(* IEC 61131-3 sources: 2026_Projet_YGO_ExcavatriceDragage/TOOLS/TEST_AUTO_CI/RESULTS/L_SIMULATION/tests (part 10) *)

TEST 'TC-T418-INT-009 Reference etablie N1 puis cycle sans depart homing'
nx := 5000; ny := 5000; raw1 := 0; raw2 := 0; previousButton := FALSE; buttonEdges := 0;
bench.Enable := TRUE; joy.Enable := TRUE; joy.ArmingPermit := TRUE; diagOk.Operational := TRUE; joy.BusCanOpenOP := diagOk; joy.JoystickOP := diagOk;
home.Enable := TRUE; home.BootReady := TRUE; home.Mode := E_Mode.MAINT_N1; home.WinchesMechanicallyStopped := TRUE;
(* Fixture deja referencee : les preuves du preset manuel reel sont dans la CI codeurs/benne et le routage PRG inchange. *)
home.M1Status.HomedAndReliable := TRUE; home.M2Status.HomedAndReliable := TRUE; home.BucketOffsetValid := TRUE;
ADVANCE_TIME(10000000); bench(RawPosM1 := raw1, RawPosM2 := raw2);
joy(RawX := bench.Operator.JoyXRaw_ANA1, RawY := bench.Operator.JoyYRaw_ANA2, RawButton := bench.Operator.JoyBtnRaw, Cfg := cfg, NeutralXMem := nx, NeutralYMem := ny);
home(DeadmanArmed := joy.DeadmanArmed, JoystickDeflected := NOT joy.AtNeutralXY, JoystickPull := joy.AxisCmdY.DirectionPositive, JoystickPush := joy.AxisCmdY.DirectionNegative, BtnValidation := bench.Operator.JoyBtnRaw);
ASSERT_EQ(home.MachineHomingSeqStep, E_MachineHomingTxState.HX0_REPOS, 'N1/cycle : aucun HX1 par geste joystick'); ASSERT_FALSE(home.M3Locked, 'N1/cycle : aucun verrou homing parasite'); ASSERT_TRUE(home.MachineHomed, 'Reference conservee');
bench.SimJoystickFwd_Up_Close_Active := TRUE;
ADVANCE_TIME(10000000); bench(RawPosM1 := raw1, RawPosM2 := raw2);
joy(RawX := bench.Operator.JoyXRaw_ANA1, RawY := bench.Operator.JoyYRaw_ANA2, RawButton := bench.Operator.JoyBtnRaw, Cfg := cfg, NeutralXMem := nx, NeutralYMem := ny);
home(DeadmanArmed := joy.DeadmanArmed, JoystickDeflected := NOT joy.AtNeutralXY, JoystickPull := joy.AxisCmdY.DirectionPositive, JoystickPush := joy.AxisCmdY.DirectionNegative, BtnValidation := bench.Operator.JoyBtnRaw);
ASSERT_EQ(home.MachineHomingSeqStep, E_MachineHomingTxState.HX0_REPOS, 'N1/cycle : aucun HX1 par geste joystick'); ASSERT_FALSE(home.M3Locked, 'N1/cycle : aucun verrou homing parasite'); ASSERT_TRUE(home.MachineHomed, 'Reference conservee');
ADVANCE_TIME(10000000); bench(RawPosM1 := raw1, RawPosM2 := raw2);
joy(RawX := bench.Operator.JoyXRaw_ANA1, RawY := bench.Operator.JoyYRaw_ANA2, RawButton := bench.Operator.JoyBtnRaw, Cfg := cfg, NeutralXMem := nx, NeutralYMem := ny);
home(DeadmanArmed := joy.DeadmanArmed, JoystickDeflected := NOT joy.AtNeutralXY, JoystickPull := joy.AxisCmdY.DirectionPositive, JoystickPush := joy.AxisCmdY.DirectionNegative, BtnValidation := bench.Operator.JoyBtnRaw);
ASSERT_EQ(home.MachineHomingSeqStep, E_MachineHomingTxState.HX0_REPOS, 'N1/cycle : aucun HX1 par geste joystick'); ASSERT_FALSE(home.M3Locked, 'N1/cycle : aucun verrou homing parasite'); ASSERT_TRUE(home.MachineHomed, 'Reference conservee');
ADVANCE_TIME(10000000); bench(RawPosM1 := raw1, RawPosM2 := raw2);
joy(RawX := bench.Operator.JoyXRaw_ANA1, RawY := bench.Operator.JoyYRaw_ANA2, RawButton := bench.Operator.JoyBtnRaw, Cfg := cfg, NeutralXMem := nx, NeutralYMem := ny);
home(DeadmanArmed := joy.DeadmanArmed, JoystickDeflected := NOT joy.AtNeutralXY, JoystickPull := joy.AxisCmdY.DirectionPositive, JoystickPush := joy.AxisCmdY.DirectionNegative, BtnValidation := bench.Operator.JoyBtnRaw);
ASSERT_EQ(home.MachineHomingSeqStep, E_MachineHomingTxState.HX0_REPOS, 'N1/cycle : aucun HX1 par geste joystick'); ASSERT_FALSE(home.M3Locked, 'N1/cycle : aucun verrou homing parasite'); ASSERT_TRUE(home.MachineHomed, 'Reference conservee');
ADVANCE_TIME(10000000); bench(RawPosM1 := raw1, RawPosM2 := raw2);
joy(RawX := bench.Operator.JoyXRaw_ANA1, RawY := bench.Operator.JoyYRaw_ANA2, RawButton := bench.Operator.JoyBtnRaw, Cfg := cfg, NeutralXMem := nx, NeutralYMem := ny);
home(DeadmanArmed := joy.DeadmanArmed, JoystickDeflected := NOT joy.AtNeutralXY, JoystickPull := joy.AxisCmdY.DirectionPositive, JoystickPush := joy.AxisCmdY.DirectionNegative, BtnValidation := bench.Operator.JoyBtnRaw);
ASSERT_EQ(home.MachineHomingSeqStep, E_MachineHomingTxState.HX0_REPOS, 'N1/cycle : aucun HX1 par geste joystick'); ASSERT_FALSE(home.M3Locked, 'N1/cycle : aucun verrou homing parasite'); ASSERT_TRUE(home.MachineHomed, 'Reference conservee');
ADVANCE_TIME(10000000); bench(RawPosM1 := raw1, RawPosM2 := raw2);
joy(RawX := bench.Operator.JoyXRaw_ANA1, RawY := bench.Operator.JoyYRaw_ANA2, RawButton := bench.Operator.JoyBtnRaw, Cfg := cfg, NeutralXMem := nx, NeutralYMem := ny);
home(DeadmanArmed := joy.DeadmanArmed, JoystickDeflected := NOT joy.AtNeutralXY, JoystickPull := joy.AxisCmdY.DirectionPositive, JoystickPush := joy.AxisCmdY.DirectionNegative, BtnValidation := bench.Operator.JoyBtnRaw);
ASSERT_EQ(home.MachineHomingSeqStep, E_MachineHomingTxState.HX0_REPOS, 'N1/cycle : aucun HX1 par geste joystick'); ASSERT_FALSE(home.M3Locked, 'N1/cycle : aucun verrou homing parasite'); ASSERT_TRUE(home.MachineHomed, 'Reference conservee');
ADVANCE_TIME(10000000); bench(RawPosM1 := raw1, RawPosM2 := raw2);
joy(RawX := bench.Operator.JoyXRaw_ANA1, RawY := bench.Operator.JoyYRaw_ANA2, RawButton := bench.Operator.JoyBtnRaw, Cfg := cfg, NeutralXMem := nx, NeutralYMem := ny);
home(DeadmanArmed := joy.DeadmanArmed, JoystickDeflected := NOT joy.AtNeutralXY, JoystickPull := joy.AxisCmdY.DirectionPositive, JoystickPush := joy.AxisCmdY.DirectionNegative, BtnValidation := bench.Operator.JoyBtnRaw);
ASSERT_EQ(home.MachineHomingSeqStep, E_MachineHomingTxState.HX0_REPOS, 'N1/cycle : aucun HX1 par geste joystick'); ASSERT_FALSE(home.M3Locked, 'N1/cycle : aucun verrou homing parasite'); ASSERT_TRUE(home.MachineHomed, 'Reference conservee');
ADVANCE_TIME(10000000); bench(RawPosM1 := raw1, RawPosM2 := raw2);
joy(RawX := bench.Operator.JoyXRaw_ANA1, RawY := bench.Operator.JoyYRaw_ANA2, RawButton := bench.Operator.JoyBtnRaw, Cfg := cfg, NeutralXMem := nx, NeutralYMem := ny);
home(DeadmanArmed := joy.DeadmanArmed, JoystickDeflected := NOT joy.AtNeutralXY, JoystickPull := joy.AxisCmdY.DirectionPositive, JoystickPush := joy.AxisCmdY.DirectionNegative, BtnValidation := bench.Operator.JoyBtnRaw);
ASSERT_EQ(home.MachineHomingSeqStep, E_MachineHomingTxState.HX0_REPOS, 'N1/cycle : aucun HX1 par geste joystick'); ASSERT_FALSE(home.M3Locked, 'N1/cycle : aucun verrou homing parasite'); ASSERT_TRUE(home.MachineHomed, 'Reference conservee');
ADVANCE_TIME(10000000); bench(RawPosM1 := raw1, RawPosM2 := raw2);
joy(RawX := bench.Operator.JoyXRaw_ANA1, RawY := bench.Operator.JoyYRaw_ANA2, RawButton := bench.Operator.JoyBtnRaw, Cfg := cfg, NeutralXMem := nx, NeutralYMem := ny);
home(DeadmanArmed := joy.DeadmanArmed, JoystickDeflected := NOT joy.AtNeutralXY, JoystickPull := joy.AxisCmdY.DirectionPositive, JoystickPush := joy.AxisCmdY.DirectionNegative, BtnValidation := bench.Operator.JoyBtnRaw);
ASSERT_EQ(home.MachineHomingSeqStep, E_MachineHomingTxState.HX0_REPOS, 'N1/cycle : aucun HX1 par geste joystick'); ASSERT_FALSE(home.M3Locked, 'N1/cycle : aucun verrou homing parasite'); ASSERT_TRUE(home.MachineHomed, 'Reference conservee');
ADVANCE_TIME(10000000); bench(RawPosM1 := raw1, RawPosM2 := raw2);
joy(RawX := bench.Operator.JoyXRaw_ANA1, RawY := bench.Operator.JoyYRaw_ANA2, RawButton := bench.Operator.JoyBtnRaw, Cfg := cfg, NeutralXMem := nx, NeutralYMem := ny);
home(DeadmanArmed := joy.DeadmanArmed, JoystickDeflected := NOT joy.AtNeutralXY, JoystickPull := joy.AxisCmdY.DirectionPositive, JoystickPush := joy.AxisCmdY.DirectionNegative, BtnValidation := bench.Operator.JoyBtnRaw);
ASSERT_EQ(home.MachineHomingSeqStep, E_MachineHomingTxState.HX0_REPOS, 'N1/cycle : aucun HX1 par geste joystick'); ASSERT_FALSE(home.M3Locked, 'N1/cycle : aucun verrou homing parasite'); ASSERT_TRUE(home.MachineHomed, 'Reference conservee');
ADVANCE_TIME(10000000); bench(RawPosM1 := raw1, RawPosM2 := raw2);
joy(RawX := bench.Operator.JoyXRaw_ANA1, RawY := bench.Operator.JoyYRaw_ANA2, RawButton := bench.Operator.JoyBtnRaw, Cfg := cfg, NeutralXMem := nx, NeutralYMem := ny);
home(DeadmanArmed := joy.DeadmanArmed, JoystickDeflected := NOT joy.AtNeutralXY, JoystickPull := joy.AxisCmdY.DirectionPositive, JoystickPush := joy.AxisCmdY.DirectionNegative, BtnValidation := bench.Operator.JoyBtnRaw);
ASSERT_EQ(home.MachineHomingSeqStep, E_MachineHomingTxState.HX0_REPOS, 'N1/cycle : aucun HX1 par geste joystick'); ASSERT_FALSE(home.M3Locked, 'N1/cycle : aucun verrou homing parasite'); ASSERT_TRUE(home.MachineHomed, 'Reference conservee');
ADVANCE_TIME(10000000); bench(RawPosM1 := raw1, RawPosM2 := raw2);
joy(RawX := bench.Operator.JoyXRaw_ANA1, RawY := bench.Operator.JoyYRaw_ANA2, RawButton := bench.Operator.JoyBtnRaw, Cfg := cfg, NeutralXMem := nx, NeutralYMem := ny);
home(DeadmanArmed := joy.DeadmanArmed, JoystickDeflected := NOT joy.AtNeutralXY, JoystickPull := joy.AxisCmdY.DirectionPositive, JoystickPush := joy.AxisCmdY.DirectionNegative, BtnValidation := bench.Operator.JoyBtnRaw);
ASSERT_EQ(home.MachineHomingSeqStep, E_MachineHomingTxState.HX0_REPOS, 'N1/cycle : aucun HX1 par geste joystick'); ASSERT_FALSE(home.M3Locked, 'N1/cycle : aucun verrou homing parasite'); ASSERT_TRUE(home.MachineHomed, 'Reference conservee');
ADVANCE_TIME(10000000); bench(RawPosM1 := raw1, RawPosM2 := raw2);
joy(RawX := bench.Operator.JoyXRaw_ANA1, RawY := bench.Operator.JoyYRaw_ANA2, RawButton := bench.Operator.JoyBtnRaw, Cfg := cfg, NeutralXMem := nx, NeutralYMem := ny);
home(DeadmanArmed := joy.DeadmanArmed, JoystickDeflected := NOT joy.AtNeutralXY, JoystickPull := joy.AxisCmdY.DirectionPositive, JoystickPush := joy.AxisCmdY.DirectionNegative, BtnValidation := bench.Operator.JoyBtnRaw);
ASSERT_EQ(home.MachineHomingSeqStep, E_MachineHomingTxState.HX0_REPOS, 'N1/cycle : aucun HX1 par geste joystick'); ASSERT_FALSE(home.M3Locked, 'N1/cycle : aucun verrou homing parasite'); ASSERT_TRUE(home.MachineHomed, 'Reference conservee');
ADVANCE_TIME(10000000); bench(RawPosM1 := raw1, RawPosM2 := raw2);
joy(RawX := bench.Operator.JoyXRaw_ANA1, RawY := bench.Operator.JoyYRaw_ANA2, RawButton := bench.Operator.JoyBtnRaw, Cfg := cfg, NeutralXMem := nx, NeutralYMem := ny);
home(DeadmanArmed := joy.DeadmanArmed, JoystickDeflected := NOT joy.AtNeutralXY, JoystickPull := joy.AxisCmdY.DirectionPositive, JoystickPush := joy.AxisCmdY.DirectionNegative, BtnValidation := bench.Operator.JoyBtnRaw);
ASSERT_EQ(home.MachineHomingSeqStep, E_MachineHomingTxState.HX0_REPOS, 'N1/cycle : aucun HX1 par geste joystick'); ASSERT_FALSE(home.M3Locked, 'N1/cycle : aucun verrou homing parasite'); ASSERT_TRUE(home.MachineHomed, 'Reference conservee');
ADVANCE_TIME(10000000); bench(RawPosM1 := raw1, RawPosM2 := raw2);
joy(RawX := bench.Operator.JoyXRaw_ANA1, RawY := bench.Operator.JoyYRaw_ANA2, RawButton := bench.Operator.JoyBtnRaw, Cfg := cfg, NeutralXMem := nx, NeutralYMem := ny);
home(DeadmanArmed := joy.DeadmanArmed, JoystickDeflected := NOT joy.AtNeutralXY, JoystickPull := joy.AxisCmdY.DirectionPositive, JoystickPush := joy.AxisCmdY.DirectionNegative, BtnValidation := bench.Operator.JoyBtnRaw);
ASSERT_EQ(home.MachineHomingSeqStep, E_MachineHomingTxState.HX0_REPOS, 'N1/cycle : aucun HX1 par geste joystick'); ASSERT_FALSE(home.M3Locked, 'N1/cycle : aucun verrou homing parasite'); ASSERT_TRUE(home.MachineHomed, 'Reference conservee');
ADVANCE_TIME(10000000); bench(RawPosM1 := raw1, RawPosM2 := raw2);
joy(RawX := bench.Operator.JoyXRaw_ANA1, RawY := bench.Operator.JoyYRaw_ANA2, RawButton := bench.Operator.JoyBtnRaw, Cfg := cfg, NeutralXMem := nx, NeutralYMem := ny);
home(DeadmanArmed := joy.DeadmanArmed, JoystickDeflected := NOT joy.AtNeutralXY, JoystickPull := joy.AxisCmdY.DirectionPositive, JoystickPush := joy.AxisCmdY.DirectionNegative, BtnValidation := bench.Operator.JoyBtnRaw);
ASSERT_EQ(home.MachineHomingSeqStep, E_MachineHomingTxState.HX0_REPOS, 'N1/cycle : aucun HX1 par geste joystick'); ASSERT_FALSE(home.M3Locked, 'N1/cycle : aucun verrou homing parasite'); ASSERT_TRUE(home.MachineHomed, 'Reference conservee');
ADVANCE_TIME(10000000); bench(RawPosM1 := raw1, RawPosM2 := raw2);
joy(RawX := bench.Operator.JoyXRaw_ANA1, RawY := bench.Operator.JoyYRaw_ANA2, RawButton := bench.Operator.JoyBtnRaw, Cfg := cfg, NeutralXMem := nx, NeutralYMem := ny);
home(DeadmanArmed := joy.DeadmanArmed, JoystickDeflected := NOT joy.AtNeutralXY, JoystickPull := joy.AxisCmdY.DirectionPositive, JoystickPush := joy.AxisCmdY.DirectionNegative, BtnValidation := bench.Operator.JoyBtnRaw);
ASSERT_EQ(home.MachineHomingSeqStep, E_MachineHomingTxState.HX0_REPOS, 'N1/cycle : aucun HX1 par geste joystick'); ASSERT_FALSE(home.M3Locked, 'N1/cycle : aucun verrou homing parasite'); ASSERT_TRUE(home.MachineHomed, 'Reference conservee');
ADVANCE_TIME(10000000); bench(RawPosM1 := raw1, RawPosM2 := raw2);
joy(RawX := bench.Operator.JoyXRaw_ANA1, RawY := bench.Operator.JoyYRaw_ANA2, RawButton := bench.Operator.JoyBtnRaw, Cfg := cfg, NeutralXMem := nx, NeutralYMem := ny);
home(DeadmanArmed := joy.DeadmanArmed, JoystickDeflected := NOT joy.AtNeutralXY, JoystickPull := joy.AxisCmdY.DirectionPositive, JoystickPush := joy.AxisCmdY.DirectionNegative, BtnValidation := bench.Operator.JoyBtnRaw);
ASSERT_EQ(home.MachineHomingSeqStep, E_MachineHomingTxState.HX0_REPOS, 'N1/cycle : aucun HX1 par geste joystick'); ASSERT_FALSE(home.M3Locked, 'N1/cycle : aucun verrou homing parasite'); ASSERT_TRUE(home.MachineHomed, 'Reference conservee');
ADVANCE_TIME(10000000); bench(RawPosM1 := raw1, RawPosM2 := raw2);
joy(RawX := bench.Operator.JoyXRaw_ANA1, RawY := bench.Operator.JoyYRaw_ANA2, RawButton := bench.Operator.JoyBtnRaw, Cfg := cfg, NeutralXMem := nx, NeutralYMem := ny);
home(DeadmanArmed := joy.DeadmanArmed, JoystickDeflected := NOT joy.AtNeutralXY, JoystickPull := joy.AxisCmdY.DirectionPositive, JoystickPush := joy.AxisCmdY.DirectionNegative, BtnValidation := bench.Operator.JoyBtnRaw);
ASSERT_EQ(home.MachineHomingSeqStep, E_MachineHomingTxState.HX0_REPOS, 'N1/cycle : aucun HX1 par geste joystick'); ASSERT_FALSE(home.M3Locked, 'N1/cycle : aucun verrou homing parasite'); ASSERT_TRUE(home.MachineHomed, 'Reference conservee');
ADVANCE_TIME(10000000); bench(RawPosM1 := raw1, RawPosM2 := raw2);
joy(RawX := bench.Operator.JoyXRaw_ANA1, RawY := bench.Operator.JoyYRaw_ANA2, RawButton := bench.Operator.JoyBtnRaw, Cfg := cfg, NeutralXMem := nx, NeutralYMem := ny);
home(DeadmanArmed := joy.DeadmanArmed, JoystickDeflected := NOT joy.AtNeutralXY, JoystickPull := joy.AxisCmdY.DirectionPositive, JoystickPush := joy.AxisCmdY.DirectionNegative, BtnValidation := bench.Operator.JoyBtnRaw);
ASSERT_EQ(home.MachineHomingSeqStep, E_MachineHomingTxState.HX0_REPOS, 'N1/cycle : aucun HX1 par geste joystick'); ASSERT_FALSE(home.M3Locked, 'N1/cycle : aucun verrou homing parasite'); ASSERT_TRUE(home.MachineHomed, 'Reference conservee');
ADVANCE_TIME(10000000); bench(RawPosM1 := raw1, RawPosM2 := raw2);
joy(RawX := bench.Operator.JoyXRaw_ANA1, RawY := bench.Operator.JoyYRaw_ANA2, RawButton := bench.Operator.JoyBtnRaw, Cfg := cfg, NeutralXMem := nx, NeutralYMem := ny);
home(DeadmanArmed := joy.DeadmanArmed, JoystickDeflected := NOT joy.AtNeutralXY, JoystickPull := joy.AxisCmdY.DirectionPositive, JoystickPush := joy.AxisCmdY.DirectionNegative, BtnValidation := bench.Operator.JoyBtnRaw);
ASSERT_EQ(home.MachineHomingSeqStep, E_MachineHomingTxState.HX0_REPOS, 'N1/cycle : aucun HX1 par geste joystick'); ASSERT_FALSE(home.M3Locked, 'N1/cycle : aucun verrou homing parasite'); ASSERT_TRUE(home.MachineHomed, 'Reference conservee');
ADVANCE_TIME(10000000); bench(RawPosM1 := raw1, RawPosM2 := raw2);
joy(RawX := bench.Operator.JoyXRaw_ANA1, RawY := bench.Operator.JoyYRaw_ANA2, RawButton := bench.Operator.JoyBtnRaw, Cfg := cfg, NeutralXMem := nx, NeutralYMem := ny);
home(DeadmanArmed := joy.DeadmanArmed, JoystickDeflected := NOT joy.AtNeutralXY, JoystickPull := joy.AxisCmdY.DirectionPositive, JoystickPush := joy.AxisCmdY.DirectionNegative, BtnValidation := bench.Operator.JoyBtnRaw);
ASSERT_EQ(home.MachineHomingSeqStep, E_MachineHomingTxState.HX0_REPOS, 'N1/cycle : aucun HX1 par geste joystick'); ASSERT_FALSE(home.M3Locked, 'N1/cycle : aucun verrou homing parasite'); ASSERT_TRUE(home.MachineHomed, 'Reference conservee');
ADVANCE_TIME(10000000); bench(RawPosM1 := raw1, RawPosM2 := raw2);
joy(RawX := bench.Operator.JoyXRaw_ANA1, RawY := bench.Operator.JoyYRaw_ANA2, RawButton := bench.Operator.JoyBtnRaw, Cfg := cfg, NeutralXMem := nx, NeutralYMem := ny);
home(DeadmanArmed := joy.DeadmanArmed, JoystickDeflected := NOT joy.AtNeutralXY, JoystickPull := joy.AxisCmdY.DirectionPositive, JoystickPush := joy.AxisCmdY.DirectionNegative, BtnValidation := bench.Operator.JoyBtnRaw);
ASSERT_EQ(home.MachineHomingSeqStep, E_MachineHomingTxState.HX0_REPOS, 'N1/cycle : aucun HX1 par geste joystick'); ASSERT_FALSE(home.M3Locked, 'N1/cycle : aucun verrou homing parasite'); ASSERT_TRUE(home.MachineHomed, 'Reference conservee');
ADVANCE_TIME(10000000); bench(RawPosM1 := raw1, RawPosM2 := raw2);
joy(RawX := bench.Operator.JoyXRaw_ANA1, RawY := bench.Operator.JoyYRaw_ANA2, RawButton := bench.Operator.JoyBtnRaw, Cfg := cfg, NeutralXMem := nx, NeutralYMem := ny);
home(DeadmanArmed := joy.DeadmanArmed, JoystickDeflected := NOT joy.AtNeutralXY, JoystickPull := joy.AxisCmdY.DirectionPositive, JoystickPush := joy.AxisCmdY.DirectionNegative, BtnValidation := bench.Operator.JoyBtnRaw);
ASSERT_EQ(home.MachineHomingSeqStep, E_MachineHomingTxState.HX0_REPOS, 'N1/cycle : aucun HX1 par geste joystick'); ASSERT_FALSE(home.M3Locked, 'N1/cycle : aucun verrou homing parasite'); ASSERT_TRUE(home.MachineHomed, 'Reference conservee');
ADVANCE_TIME(10000000); bench(RawPosM1 := raw1, RawPosM2 := raw2);
joy(RawX := bench.Operator.JoyXRaw_ANA1, RawY := bench.Operator.JoyYRaw_ANA2, RawButton := bench.Operator.JoyBtnRaw, Cfg := cfg, NeutralXMem := nx, NeutralYMem := ny);
home(DeadmanArmed := joy.DeadmanArmed, JoystickDeflected := NOT joy.AtNeutralXY, JoystickPull := joy.AxisCmdY.DirectionPositive, JoystickPush := joy.AxisCmdY.DirectionNegative, BtnValidation := bench.Operator.JoyBtnRaw);
ASSERT_EQ(home.MachineHomingSeqStep, E_MachineHomingTxState.HX0_REPOS, 'N1/cycle : aucun HX1 par geste joystick'); ASSERT_FALSE(home.M3Locked, 'N1/cycle : aucun verrou homing parasite'); ASSERT_TRUE(home.MachineHomed, 'Reference conservee');
ADVANCE_TIME(10000000); bench(RawPosM1 := raw1, RawPosM2 := raw2);
joy(RawX := bench.Operator.JoyXRaw_ANA1, RawY := bench.Operator.JoyYRaw_ANA2, RawButton := bench.Operator.JoyBtnRaw, Cfg := cfg, NeutralXMem := nx, NeutralYMem := ny);
home(DeadmanArmed := joy.DeadmanArmed, JoystickDeflected := NOT joy.AtNeutralXY, JoystickPull := joy.AxisCmdY.DirectionPositive, JoystickPush := joy.AxisCmdY.DirectionNegative, BtnValidation := bench.Operator.JoyBtnRaw);
ASSERT_EQ(home.MachineHomingSeqStep, E_MachineHomingTxState.HX0_REPOS, 'N1/cycle : aucun HX1 par geste joystick'); ASSERT_FALSE(home.M3Locked, 'N1/cycle : aucun verrou homing parasite'); ASSERT_TRUE(home.MachineHomed, 'Reference conservee');
ADVANCE_TIME(10000000); bench(RawPosM1 := raw1, RawPosM2 := raw2);
joy(RawX := bench.Operator.JoyXRaw_ANA1, RawY := bench.Operator.JoyYRaw_ANA2, RawButton := bench.Operator.JoyBtnRaw, Cfg := cfg, NeutralXMem := nx, NeutralYMem := ny);
home(DeadmanArmed := joy.DeadmanArmed, JoystickDeflected := NOT joy.AtNeutralXY, JoystickPull := joy.AxisCmdY.DirectionPositive, JoystickPush := joy.AxisCmdY.DirectionNegative, BtnValidation := bench.Operator.JoyBtnRaw);
ASSERT_EQ(home.MachineHomingSeqStep, E_MachineHomingTxState.HX0_REPOS, 'N1/cycle : aucun HX1 par geste joystick'); ASSERT_FALSE(home.M3Locked, 'N1/cycle : aucun verrou homing parasite'); ASSERT_TRUE(home.MachineHomed, 'Reference conservee');
ADVANCE_TIME(10000000); bench(RawPosM1 := raw1, RawPosM2 := raw2);
joy(RawX := bench.Operator.JoyXRaw_ANA1, RawY := bench.Operator.JoyYRaw_ANA2, RawButton := bench.Operator.JoyBtnRaw, Cfg := cfg, NeutralXMem := nx, NeutralYMem := ny);
home(DeadmanArmed := joy.DeadmanArmed, JoystickDeflected := NOT joy.AtNeutralXY, JoystickPull := joy.AxisCmdY.DirectionPositive, JoystickPush := joy.AxisCmdY.DirectionNegative, BtnValidation := bench.Operator.JoyBtnRaw);
ASSERT_EQ(home.MachineHomingSeqStep, E_MachineHomingTxState.HX0_REPOS, 'N1/cycle : aucun HX1 par geste joystick'); ASSERT_FALSE(home.M3Locked, 'N1/cycle : aucun verrou homing parasite'); ASSERT_TRUE(home.MachineHomed, 'Reference conservee');
ADVANCE_TIME(10000000); bench(RawPosM1 := raw1, RawPosM2 := raw2);
joy(RawX := bench.Operator.JoyXRaw_ANA1, RawY := bench.Operator.JoyYRaw_ANA2, RawButton := bench.Operator.JoyBtnRaw, Cfg := cfg, NeutralXMem := nx, NeutralYMem := ny);
home(DeadmanArmed := joy.DeadmanArmed, JoystickDeflected := NOT joy.AtNeutralXY, JoystickPull := joy.AxisCmdY.DirectionPositive, JoystickPush := joy.AxisCmdY.DirectionNegative, BtnValidation := bench.Operator.JoyBtnRaw);
ASSERT_EQ(home.MachineHomingSeqStep, E_MachineHomingTxState.HX0_REPOS, 'N1/cycle : aucun HX1 par geste joystick'); ASSERT_FALSE(home.M3Locked, 'N1/cycle : aucun verrou homing parasite'); ASSERT_TRUE(home.MachineHomed, 'Reference conservee');
ADVANCE_TIME(10000000); bench(RawPosM1 := raw1, RawPosM2 := raw2);
joy(RawX := bench.Operator.JoyXRaw_ANA1, RawY := bench.Operator.JoyYRaw_ANA2, RawButton := bench.Operator.JoyBtnRaw, Cfg := cfg, NeutralXMem := nx, NeutralYMem := ny);
home(DeadmanArmed := joy.DeadmanArmed, JoystickDeflected := NOT joy.AtNeutralXY, JoystickPull := joy.AxisCmdY.DirectionPositive, JoystickPush := joy.AxisCmdY.DirectionNegative, BtnValidation := bench.Operator.JoyBtnRaw);
ASSERT_EQ(home.MachineHomingSeqStep, E_MachineHomingTxState.HX0_REPOS, 'N1/cycle : aucun HX1 par geste joystick'); ASSERT_FALSE(home.M3Locked, 'N1/cycle : aucun verrou homing parasite'); ASSERT_TRUE(home.MachineHomed, 'Reference conservee');
ADVANCE_TIME(10000000); bench(RawPosM1 := raw1, RawPosM2 := raw2);
joy(RawX := bench.Operator.JoyXRaw_ANA1, RawY := bench.Operator.JoyYRaw_ANA2, RawButton := bench.Operator.JoyBtnRaw, Cfg := cfg, NeutralXMem := nx, NeutralYMem := ny);
home(DeadmanArmed := joy.DeadmanArmed, JoystickDeflected := NOT joy.AtNeutralXY, JoystickPull := joy.AxisCmdY.DirectionPositive, JoystickPush := joy.AxisCmdY.DirectionNegative, BtnValidation := bench.Operator.JoyBtnRaw);
ASSERT_EQ(home.MachineHomingSeqStep, E_MachineHomingTxState.HX0_REPOS, 'N1/cycle : aucun HX1 par geste joystick'); ASSERT_FALSE(home.M3Locked, 'N1/cycle : aucun verrou homing parasite'); ASSERT_TRUE(home.MachineHomed, 'Reference conservee');
ADVANCE_TIME(10000000); bench(RawPosM1 := raw1, RawPosM2 := raw2);
joy(RawX := bench.Operator.JoyXRaw_ANA1, RawY := bench.Operator.JoyYRaw_ANA2, RawButton := bench.Operator.JoyBtnRaw, Cfg := cfg, NeutralXMem := nx, NeutralYMem := ny);
home(DeadmanArmed := joy.DeadmanArmed, JoystickDeflected := NOT joy.AtNeutralXY, JoystickPull := joy.AxisCmdY.DirectionPositive, JoystickPush := joy.AxisCmdY.DirectionNegative, BtnValidation := bench.Operator.JoyBtnRaw);
ASSERT_EQ(home.MachineHomingSeqStep, E_MachineHomingTxState.HX0_REPOS, 'N1/cycle : aucun HX1 par geste joystick'); ASSERT_FALSE(home.M3Locked, 'N1/cycle : aucun verrou homing parasite'); ASSERT_TRUE(home.MachineHomed, 'Reference conservee');
ADVANCE_TIME(10000000); bench(RawPosM1 := raw1, RawPosM2 := raw2);
joy(RawX := bench.Operator.JoyXRaw_ANA1, RawY := bench.Operator.JoyYRaw_ANA2, RawButton := bench.Operator.JoyBtnRaw, Cfg := cfg, NeutralXMem := nx, NeutralYMem := ny);
home(DeadmanArmed := joy.DeadmanArmed, JoystickDeflected := NOT joy.AtNeutralXY, JoystickPull := joy.AxisCmdY.DirectionPositive, JoystickPush := joy.AxisCmdY.DirectionNegative, BtnValidation := bench.Operator.JoyBtnRaw);
ASSERT_EQ(home.MachineHomingSeqStep, E_MachineHomingTxState.HX0_REPOS, 'N1/cycle : aucun HX1 par geste joystick'); ASSERT_FALSE(home.M3Locked, 'N1/cycle : aucun verrou homing parasite'); ASSERT_TRUE(home.MachineHomed, 'Reference conservee');
ADVANCE_TIME(10000000); bench(RawPosM1 := raw1, RawPosM2 := raw2);
joy(RawX := bench.Operator.JoyXRaw_ANA1, RawY := bench.Operator.JoyYRaw_ANA2, RawButton := bench.Operator.JoyBtnRaw, Cfg := cfg, NeutralXMem := nx, NeutralYMem := ny);
home(DeadmanArmed := joy.DeadmanArmed, JoystickDeflected := NOT joy.AtNeutralXY, JoystickPull := joy.AxisCmdY.DirectionPositive, JoystickPush := joy.AxisCmdY.DirectionNegative, BtnValidation := bench.Operator.JoyBtnRaw);
ASSERT_EQ(home.MachineHomingSeqStep, E_MachineHomingTxState.HX0_REPOS, 'N1/cycle : aucun HX1 par geste joystick'); ASSERT_FALSE(home.M3Locked, 'N1/cycle : aucun verrou homing parasite'); ASSERT_TRUE(home.MachineHomed, 'Reference conservee');
ADVANCE_TIME(10000000); bench(RawPosM1 := raw1, RawPosM2 := raw2);
joy(RawX := bench.Operator.JoyXRaw_ANA1, RawY := bench.Operator.JoyYRaw_ANA2, RawButton := bench.Operator.JoyBtnRaw, Cfg := cfg, NeutralXMem := nx, NeutralYMem := ny);
home(DeadmanArmed := joy.DeadmanArmed, JoystickDeflected := NOT joy.AtNeutralXY, JoystickPull := joy.AxisCmdY.DirectionPositive, JoystickPush := joy.AxisCmdY.DirectionNegative, BtnValidation := bench.Operator.JoyBtnRaw);
ASSERT_EQ(home.MachineHomingSeqStep, E_MachineHomingTxState.HX0_REPOS, 'N1/cycle : aucun HX1 par geste joystick'); ASSERT_FALSE(home.M3Locked, 'N1/cycle : aucun verrou homing parasite'); ASSERT_TRUE(home.MachineHomed, 'Reference conservee');
ADVANCE_TIME(10000000); bench(RawPosM1 := raw1, RawPosM2 := raw2);
joy(RawX := bench.Operator.JoyXRaw_ANA1, RawY := bench.Operator.JoyYRaw_ANA2, RawButton := bench.Operator.JoyBtnRaw, Cfg := cfg, NeutralXMem := nx, NeutralYMem := ny);
home(DeadmanArmed := joy.DeadmanArmed, JoystickDeflected := NOT joy.AtNeutralXY, JoystickPull := joy.AxisCmdY.DirectionPositive, JoystickPush := joy.AxisCmdY.DirectionNegative, BtnValidation := bench.Operator.JoyBtnRaw);
ASSERT_EQ(home.MachineHomingSeqStep, E_MachineHomingTxState.HX0_REPOS, 'N1/cycle : aucun HX1 par geste joystick'); ASSERT_FALSE(home.M3Locked, 'N1/cycle : aucun verrou homing parasite'); ASSERT_TRUE(home.MachineHomed, 'Reference conservee');
ADVANCE_TIME(10000000); bench(RawPosM1 := raw1, RawPosM2 := raw2);
joy(RawX := bench.Operator.JoyXRaw_ANA1, RawY := bench.Operator.JoyYRaw_ANA2, RawButton := bench.Operator.JoyBtnRaw, Cfg := cfg, NeutralXMem := nx, NeutralYMem := ny);
home(DeadmanArmed := joy.DeadmanArmed, JoystickDeflected := NOT joy.AtNeutralXY, JoystickPull := joy.AxisCmdY.DirectionPositive, JoystickPush := joy.AxisCmdY.DirectionNegative, BtnValidation := bench.Operator.JoyBtnRaw);
ASSERT_EQ(home.MachineHomingSeqStep, E_MachineHomingTxState.HX0_REPOS, 'N1/cycle : aucun HX1 par geste joystick'); ASSERT_FALSE(home.M3Locked, 'N1/cycle : aucun verrou homing parasite'); ASSERT_TRUE(home.MachineHomed, 'Reference conservee');
ADVANCE_TIME(10000000); bench(RawPosM1 := raw1, RawPosM2 := raw2);
joy(RawX := bench.Operator.JoyXRaw_ANA1, RawY := bench.Operator.JoyYRaw_ANA2, RawButton := bench.Operator.JoyBtnRaw, Cfg := cfg, NeutralXMem := nx, NeutralYMem := ny);
home(DeadmanArmed := joy.DeadmanArmed, JoystickDeflected := NOT joy.AtNeutralXY, JoystickPull := joy.AxisCmdY.DirectionPositive, JoystickPush := joy.AxisCmdY.DirectionNegative, BtnValidation := bench.Operator.JoyBtnRaw);
ASSERT_EQ(home.MachineHomingSeqStep, E_MachineHomingTxState.HX0_REPOS, 'N1/cycle : aucun HX1 par geste joystick'); ASSERT_FALSE(home.M3Locked, 'N1/cycle : aucun verrou homing parasite'); ASSERT_TRUE(home.MachineHomed, 'Reference conservee');
ADVANCE_TIME(10000000); bench(RawPosM1 := raw1, RawPosM2 := raw2);
joy(RawX := bench.Operator.JoyXRaw_ANA1, RawY := bench.Operator.JoyYRaw_ANA2, RawButton := bench.Operator.JoyBtnRaw, Cfg := cfg, NeutralXMem := nx, NeutralYMem := ny);
home(DeadmanArmed := joy.DeadmanArmed, JoystickDeflected := NOT joy.AtNeutralXY, JoystickPull := joy.AxisCmdY.DirectionPositive, JoystickPush := joy.AxisCmdY.DirectionNegative, BtnValidation := bench.Operator.JoyBtnRaw);
ASSERT_EQ(home.MachineHomingSeqStep, E_MachineHomingTxState.HX0_REPOS, 'N1/cycle : aucun HX1 par geste joystick'); ASSERT_FALSE(home.M3Locked, 'N1/cycle : aucun verrou homing parasite'); ASSERT_TRUE(home.MachineHomed, 'Reference conservee');
ADVANCE_TIME(10000000); bench(RawPosM1 := raw1, RawPosM2 := raw2);
joy(RawX := bench.Operator.JoyXRaw_ANA1, RawY := bench.Operator.JoyYRaw_ANA2, RawButton := bench.Operator.JoyBtnRaw, Cfg := cfg, NeutralXMem := nx, NeutralYMem := ny);
home(DeadmanArmed := joy.DeadmanArmed, JoystickDeflected := NOT joy.AtNeutralXY, JoystickPull := joy.AxisCmdY.DirectionPositive, JoystickPush := joy.AxisCmdY.DirectionNegative, BtnValidation := bench.Operator.JoyBtnRaw);
ASSERT_EQ(home.MachineHomingSeqStep, E_MachineHomingTxState.HX0_REPOS, 'N1/cycle : aucun HX1 par geste joystick'); ASSERT_FALSE(home.M3Locked, 'N1/cycle : aucun verrou homing parasite'); ASSERT_TRUE(home.MachineHomed, 'Reference conservee');
ADVANCE_TIME(10000000); bench(RawPosM1 := raw1, RawPosM2 := raw2);
joy(RawX := bench.Operator.JoyXRaw_ANA1, RawY := bench.Operator.JoyYRaw_ANA2, RawButton := bench.Operator.JoyBtnRaw, Cfg := cfg, NeutralXMem := nx, NeutralYMem := ny);
home(DeadmanArmed := joy.DeadmanArmed, JoystickDeflected := NOT joy.AtNeutralXY, JoystickPull := joy.AxisCmdY.DirectionPositive, JoystickPush := joy.AxisCmdY.DirectionNegative, BtnValidation := bench.Operator.JoyBtnRaw);
ASSERT_EQ(home.MachineHomingSeqStep, E_MachineHomingTxState.HX0_REPOS, 'N1/cycle : aucun HX1 par geste joystick'); ASSERT_FALSE(home.M3Locked, 'N1/cycle : aucun verrou homing parasite'); ASSERT_TRUE(home.MachineHomed, 'Reference conservee');
ADVANCE_TIME(10000000); bench(RawPosM1 := raw1, RawPosM2 := raw2);
joy(RawX := bench.Operator.JoyXRaw_ANA1, RawY := bench.Operator.JoyYRaw_ANA2, RawButton := bench.Operator.JoyBtnRaw, Cfg := cfg, NeutralXMem := nx, NeutralYMem := ny);
home(DeadmanArmed := joy.DeadmanArmed, JoystickDeflected := NOT joy.AtNeutralXY, JoystickPull := joy.AxisCmdY.DirectionPositive, JoystickPush := joy.AxisCmdY.DirectionNegative, BtnValidation := bench.Operator.JoyBtnRaw);
ASSERT_EQ(home.MachineHomingSeqStep, E_MachineHomingTxState.HX0_REPOS, 'N1/cycle : aucun HX1 par geste joystick'); ASSERT_FALSE(home.M3Locked, 'N1/cycle : aucun verrou homing parasite'); ASSERT_TRUE(home.MachineHomed, 'Reference conservee');
ADVANCE_TIME(10000000); bench(RawPosM1 := raw1, RawPosM2 := raw2);
joy(RawX := bench.Operator.JoyXRaw_ANA1, RawY := bench.Operator.JoyYRaw_ANA2, RawButton := bench.Operator.JoyBtnRaw, Cfg := cfg, NeutralXMem := nx, NeutralYMem := ny);
home(DeadmanArmed := joy.DeadmanArmed, JoystickDeflected := NOT joy.AtNeutralXY, JoystickPull := joy.AxisCmdY.DirectionPositive, JoystickPush := joy.AxisCmdY.DirectionNegative, BtnValidation := bench.Operator.JoyBtnRaw);
ASSERT_EQ(home.MachineHomingSeqStep, E_MachineHomingTxState.HX0_REPOS, 'N1/cycle : aucun HX1 par geste joystick'); ASSERT_FALSE(home.M3Locked, 'N1/cycle : aucun verrou homing parasite'); ASSERT_TRUE(home.MachineHomed, 'Reference conservee');
ADVANCE_TIME(10000000); bench(RawPosM1 := raw1, RawPosM2 := raw2);
joy(RawX := bench.Operator.JoyXRaw_ANA1, RawY := bench.Operator.JoyYRaw_ANA2, RawButton := bench.Operator.JoyBtnRaw, Cfg := cfg, NeutralXMem := nx, NeutralYMem := ny);
home(DeadmanArmed := joy.DeadmanArmed, JoystickDeflected := NOT joy.AtNeutralXY, JoystickPull := joy.AxisCmdY.DirectionPositive, JoystickPush := joy.AxisCmdY.DirectionNegative, BtnValidation := bench.Operator.JoyBtnRaw);
ASSERT_EQ(home.MachineHomingSeqStep, E_MachineHomingTxState.HX0_REPOS, 'N1/cycle : aucun HX1 par geste joystick'); ASSERT_FALSE(home.M3Locked, 'N1/cycle : aucun verrou homing parasite'); ASSERT_TRUE(home.MachineHomed, 'Reference conservee');
ADVANCE_TIME(10000000); bench(RawPosM1 := raw1, RawPosM2 := raw2);
joy(RawX := bench.Operator.JoyXRaw_ANA1, RawY := bench.Operator.JoyYRaw_ANA2, RawButton := bench.Operator.JoyBtnRaw, Cfg := cfg, NeutralXMem := nx, NeutralYMem := ny);
home(DeadmanArmed := joy.DeadmanArmed, JoystickDeflected := NOT joy.AtNeutralXY, JoystickPull := joy.AxisCmdY.DirectionPositive, JoystickPush := joy.AxisCmdY.DirectionNegative, BtnValidation := bench.Operator.JoyBtnRaw);
ASSERT_EQ(home.MachineHomingSeqStep, E_MachineHomingTxState.HX0_REPOS, 'N1/cycle : aucun HX1 par geste joystick'); ASSERT_FALSE(home.M3Locked, 'N1/cycle : aucun verrou homing parasite'); ASSERT_TRUE(home.MachineHomed, 'Reference conservee');
ADVANCE_TIME(10000000); bench(RawPosM1 := raw1, RawPosM2 := raw2);
joy(RawX := bench.Operator.JoyXRaw_ANA1, RawY := bench.Operator.JoyYRaw_ANA2, RawButton := bench.Operator.JoyBtnRaw, Cfg := cfg, NeutralXMem := nx, NeutralYMem := ny);
home(DeadmanArmed := joy.DeadmanArmed, JoystickDeflected := NOT joy.AtNeutralXY, JoystickPull := joy.AxisCmdY.DirectionPositive, JoystickPush := joy.AxisCmdY.DirectionNegative, BtnValidation := bench.Operator.JoyBtnRaw);
ASSERT_EQ(home.MachineHomingSeqStep, E_MachineHomingTxState.HX0_REPOS, 'N1/cycle : aucun HX1 par geste joystick'); ASSERT_FALSE(home.M3Locked, 'N1/cycle : aucun verrou homing parasite'); ASSERT_TRUE(home.MachineHomed, 'Reference conservee');
ADVANCE_TIME(10000000); bench(RawPosM1 := raw1, RawPosM2 := raw2);
joy(RawX := bench.Operator.JoyXRaw_ANA1, RawY := bench.Operator.JoyYRaw_ANA2, RawButton := bench.Operator.JoyBtnRaw, Cfg := cfg, NeutralXMem := nx, NeutralYMem := ny);
home(DeadmanArmed := joy.DeadmanArmed, JoystickDeflected := NOT joy.AtNeutralXY, JoystickPull := joy.AxisCmdY.DirectionPositive, JoystickPush := joy.AxisCmdY.DirectionNegative, BtnValidation := bench.Operator.JoyBtnRaw);
ASSERT_EQ(home.MachineHomingSeqStep, E_MachineHomingTxState.HX0_REPOS, 'N1/cycle : aucun HX1 par geste joystick'); ASSERT_FALSE(home.M3Locked, 'N1/cycle : aucun verrou homing parasite'); ASSERT_TRUE(home.MachineHomed, 'Reference conservee');
ADVANCE_TIME(10000000); bench(RawPosM1 := raw1, RawPosM2 := raw2);
joy(RawX := bench.Operator.JoyXRaw_ANA1, RawY := bench.Operator.JoyYRaw_ANA2, RawButton := bench.Operator.JoyBtnRaw, Cfg := cfg, NeutralXMem := nx, NeutralYMem := ny);
home(DeadmanArmed := joy.DeadmanArmed, JoystickDeflected := NOT joy.AtNeutralXY, JoystickPull := joy.AxisCmdY.DirectionPositive, JoystickPush := joy.AxisCmdY.DirectionNegative, BtnValidation := bench.Operator.JoyBtnRaw);
ASSERT_EQ(home.MachineHomingSeqStep, E_MachineHomingTxState.HX0_REPOS, 'N1/cycle : aucun HX1 par geste joystick'); ASSERT_FALSE(home.M3Locked, 'N1/cycle : aucun verrou homing parasite'); ASSERT_TRUE(home.MachineHomed, 'Reference conservee');
ADVANCE_TIME(10000000); bench(RawPosM1 := raw1, RawPosM2 := raw2);
joy(RawX := bench.Operator.JoyXRaw_ANA1, RawY := bench.Operator.JoyYRaw_ANA2, RawButton := bench.Operator.JoyBtnRaw, Cfg := cfg, NeutralXMem := nx, NeutralYMem := ny);
home(DeadmanArmed := joy.DeadmanArmed, JoystickDeflected := NOT joy.AtNeutralXY, JoystickPull := joy.AxisCmdY.DirectionPositive, JoystickPush := joy.AxisCmdY.DirectionNegative, BtnValidation := bench.Operator.JoyBtnRaw);
ASSERT_EQ(home.MachineHomingSeqStep, E_MachineHomingTxState.HX0_REPOS, 'N1/cycle : aucun HX1 par geste joystick'); ASSERT_FALSE(home.M3Locked, 'N1/cycle : aucun verrou homing parasite'); ASSERT_TRUE(home.MachineHomed, 'Reference conservee');
ADVANCE_TIME(10000000); bench(RawPosM1 := raw1, RawPosM2 := raw2);
joy(RawX := bench.Operator.JoyXRaw_ANA1, RawY := bench.Operator.JoyYRaw_ANA2, RawButton := bench.Operator.JoyBtnRaw, Cfg := cfg, NeutralXMem := nx, NeutralYMem := ny);
home(DeadmanArmed := joy.DeadmanArmed, JoystickDeflected := NOT joy.AtNeutralXY, JoystickPull := joy.AxisCmdY.DirectionPositive, JoystickPush := joy.AxisCmdY.DirectionNegative, BtnValidation := bench.Operator.JoyBtnRaw);
ASSERT_EQ(home.MachineHomingSeqStep, E_MachineHomingTxState.HX0_REPOS, 'N1/cycle : aucun HX1 par geste joystick'); ASSERT_FALSE(home.M3Locked, 'N1/cycle : aucun verrou homing parasite'); ASSERT_TRUE(home.MachineHomed, 'Reference conservee');
ADVANCE_TIME(10000000); bench(RawPosM1 := raw1, RawPosM2 := raw2);
joy(RawX := bench.Operator.JoyXRaw_ANA1, RawY := bench.Operator.JoyYRaw_ANA2, RawButton := bench.Operator.JoyBtnRaw, Cfg := cfg, NeutralXMem := nx, NeutralYMem := ny);
home(DeadmanArmed := joy.DeadmanArmed, JoystickDeflected := NOT joy.AtNeutralXY, JoystickPull := joy.AxisCmdY.DirectionPositive, JoystickPush := joy.AxisCmdY.DirectionNegative, BtnValidation := bench.Operator.JoyBtnRaw);
ASSERT_EQ(home.MachineHomingSeqStep, E_MachineHomingTxState.HX0_REPOS, 'N1/cycle : aucun HX1 par geste joystick'); ASSERT_FALSE(home.M3Locked, 'N1/cycle : aucun verrou homing parasite'); ASSERT_TRUE(home.MachineHomed, 'Reference conservee');
ADVANCE_TIME(10000000); bench(RawPosM1 := raw1, RawPosM2 := raw2);
joy(RawX := bench.Operator.JoyXRaw_ANA1, RawY := bench.Operator.JoyYRaw_ANA2, RawButton := bench.Operator.JoyBtnRaw, Cfg := cfg, NeutralXMem := nx, NeutralYMem := ny);
home(DeadmanArmed := joy.DeadmanArmed, JoystickDeflected := NOT joy.AtNeutralXY, JoystickPull := joy.AxisCmdY.DirectionPositive, JoystickPush := joy.AxisCmdY.DirectionNegative, BtnValidation := bench.Operator.JoyBtnRaw);
ASSERT_EQ(home.MachineHomingSeqStep, E_MachineHomingTxState.HX0_REPOS, 'N1/cycle : aucun HX1 par geste joystick'); ASSERT_FALSE(home.M3Locked, 'N1/cycle : aucun verrou homing parasite'); ASSERT_TRUE(home.MachineHomed, 'Reference conservee');
ADVANCE_TIME(10000000); bench(RawPosM1 := raw1, RawPosM2 := raw2);
joy(RawX := bench.Operator.JoyXRaw_ANA1, RawY := bench.Operator.JoyYRaw_ANA2, RawButton := bench.Operator.JoyBtnRaw, Cfg := cfg, NeutralXMem := nx, NeutralYMem := ny);
home(DeadmanArmed := joy.DeadmanArmed, JoystickDeflected := NOT joy.AtNeutralXY, JoystickPull := joy.AxisCmdY.DirectionPositive, JoystickPush := joy.AxisCmdY.DirectionNegative, BtnValidation := bench.Operator.JoyBtnRaw);
ASSERT_EQ(home.MachineHomingSeqStep, E_MachineHomingTxState.HX0_REPOS, 'N1/cycle : aucun HX1 par geste joystick'); ASSERT_FALSE(home.M3Locked, 'N1/cycle : aucun verrou homing parasite'); ASSERT_TRUE(home.MachineHomed, 'Reference conservee');
ADVANCE_TIME(10000000); bench(RawPosM1 := raw1, RawPosM2 := raw2);
joy(RawX := bench.Operator.JoyXRaw_ANA1, RawY := bench.Operator.JoyYRaw_ANA2, RawButton := bench.Operator.JoyBtnRaw, Cfg := cfg, NeutralXMem := nx, NeutralYMem := ny);
home(DeadmanArmed := joy.DeadmanArmed, JoystickDeflected := NOT joy.AtNeutralXY, JoystickPull := joy.AxisCmdY.DirectionPositive, JoystickPush := joy.AxisCmdY.DirectionNegative, BtnValidation := bench.Operator.JoyBtnRaw);
ASSERT_EQ(home.MachineHomingSeqStep, E_MachineHomingTxState.HX0_REPOS, 'N1/cycle : aucun HX1 par geste joystick'); ASSERT_FALSE(home.M3Locked, 'N1/cycle : aucun verrou homing parasite'); ASSERT_TRUE(home.MachineHomed, 'Reference conservee');
ADVANCE_TIME(10000000); bench(RawPosM1 := raw1, RawPosM2 := raw2);
joy(RawX := bench.Operator.JoyXRaw_ANA1, RawY := bench.Operator.JoyYRaw_ANA2, RawButton := bench.Operator.JoyBtnRaw, Cfg := cfg, NeutralXMem := nx, NeutralYMem := ny);
home(DeadmanArmed := joy.DeadmanArmed, JoystickDeflected := NOT joy.AtNeutralXY, JoystickPull := joy.AxisCmdY.DirectionPositive, JoystickPush := joy.AxisCmdY.DirectionNegative, BtnValidation := bench.Operator.JoyBtnRaw);
ASSERT_EQ(home.MachineHomingSeqStep, E_MachineHomingTxState.HX0_REPOS, 'N1/cycle : aucun HX1 par geste joystick'); ASSERT_FALSE(home.M3Locked, 'N1/cycle : aucun verrou homing parasite'); ASSERT_TRUE(home.MachineHomed, 'Reference conservee');
ADVANCE_TIME(10000000); bench(RawPosM1 := raw1, RawPosM2 := raw2);
joy(RawX := bench.Operator.JoyXRaw_ANA1, RawY := bench.Operator.JoyYRaw_ANA2, RawButton := bench.Operator.JoyBtnRaw, Cfg := cfg, NeutralXMem := nx, NeutralYMem := ny);
home(DeadmanArmed := joy.DeadmanArmed, JoystickDeflected := NOT joy.AtNeutralXY, JoystickPull := joy.AxisCmdY.DirectionPositive, JoystickPush := joy.AxisCmdY.DirectionNegative, BtnValidation := bench.Operator.JoyBtnRaw);
ASSERT_EQ(home.MachineHomingSeqStep, E_MachineHomingTxState.HX0_REPOS, 'N1/cycle : aucun HX1 par geste joystick'); ASSERT_FALSE(home.M3Locked, 'N1/cycle : aucun verrou homing parasite'); ASSERT_TRUE(home.MachineHomed, 'Reference conservee');
ADVANCE_TIME(10000000); bench(RawPosM1 := raw1, RawPosM2 := raw2);
joy(RawX := bench.Operator.JoyXRaw_ANA1, RawY := bench.Operator.JoyYRaw_ANA2, RawButton := bench.Operator.JoyBtnRaw, Cfg := cfg, NeutralXMem := nx, NeutralYMem := ny);
home(DeadmanArmed := joy.DeadmanArmed, JoystickDeflected := NOT joy.AtNeutralXY, JoystickPull := joy.AxisCmdY.DirectionPositive, JoystickPush := joy.AxisCmdY.DirectionNegative, BtnValidation := bench.Operator.JoyBtnRaw);
ASSERT_EQ(home.MachineHomingSeqStep, E_MachineHomingTxState.HX0_REPOS, 'N1/cycle : aucun HX1 par geste joystick'); ASSERT_FALSE(home.M3Locked, 'N1/cycle : aucun verrou homing parasite'); ASSERT_TRUE(home.MachineHomed, 'Reference conservee');
ADVANCE_TIME(10000000); bench(RawPosM1 := raw1, RawPosM2 := raw2);
joy(RawX := bench.Operator.JoyXRaw_ANA1, RawY := bench.Operator.JoyYRaw_ANA2, RawButton := bench.Operator.JoyBtnRaw, Cfg := cfg, NeutralXMem := nx, NeutralYMem := ny);
home(DeadmanArmed := joy.DeadmanArmed, JoystickDeflected := NOT joy.AtNeutralXY, JoystickPull := joy.AxisCmdY.DirectionPositive, JoystickPush := joy.AxisCmdY.DirectionNegative, BtnValidation := bench.Operator.JoyBtnRaw);
ASSERT_EQ(home.MachineHomingSeqStep, E_MachineHomingTxState.HX0_REPOS, 'N1/cycle : aucun HX1 par geste joystick'); ASSERT_FALSE(home.M3Locked, 'N1/cycle : aucun verrou homing parasite'); ASSERT_TRUE(home.MachineHomed, 'Reference conservee');
ADVANCE_TIME(10000000); bench(RawPosM1 := raw1, RawPosM2 := raw2);
joy(RawX := bench.Operator.JoyXRaw_ANA1, RawY := bench.Operator.JoyYRaw_ANA2, RawButton := bench.Operator.JoyBtnRaw, Cfg := cfg, NeutralXMem := nx, NeutralYMem := ny);
home(DeadmanArmed := joy.DeadmanArmed, JoystickDeflected := NOT joy.AtNeutralXY, JoystickPull := joy.AxisCmdY.DirectionPositive, JoystickPush := joy.AxisCmdY.DirectionNegative, BtnValidation := bench.Operator.JoyBtnRaw);
ASSERT_EQ(home.MachineHomingSeqStep, E_MachineHomingTxState.HX0_REPOS, 'N1/cycle : aucun HX1 par geste joystick'); ASSERT_FALSE(home.M3Locked, 'N1/cycle : aucun verrou homing parasite'); ASSERT_TRUE(home.MachineHomed, 'Reference conservee');
ADVANCE_TIME(10000000); bench(RawPosM1 := raw1, RawPosM2 := raw2);
joy(RawX := bench.Operator.JoyXRaw_ANA1, RawY := bench.Operator.JoyYRaw_ANA2, RawButton := bench.Operator.JoyBtnRaw, Cfg := cfg, NeutralXMem := nx, NeutralYMem := ny);
home(DeadmanArmed := joy.DeadmanArmed, JoystickDeflected := NOT joy.AtNeutralXY, JoystickPull := joy.AxisCmdY.DirectionPositive, JoystickPush := joy.AxisCmdY.DirectionNegative, BtnValidation := bench.Operator.JoyBtnRaw);
ASSERT_EQ(home.MachineHomingSeqStep, E_MachineHomingTxState.HX0_REPOS, 'N1/cycle : aucun HX1 par geste joystick'); ASSERT_FALSE(home.M3Locked, 'N1/cycle : aucun verrou homing parasite'); ASSERT_TRUE(home.MachineHomed, 'Reference conservee');
ADVANCE_TIME(10000000); bench(RawPosM1 := raw1, RawPosM2 := raw2);
joy(RawX := bench.Operator.JoyXRaw_ANA1, RawY := bench.Operator.JoyYRaw_ANA2, RawButton := bench.Operator.JoyBtnRaw, Cfg := cfg, NeutralXMem := nx, NeutralYMem := ny);
home(DeadmanArmed := joy.DeadmanArmed, JoystickDeflected := NOT joy.AtNeutralXY, JoystickPull := joy.AxisCmdY.DirectionPositive, JoystickPush := joy.AxisCmdY.DirectionNegative, BtnValidation := bench.Operator.JoyBtnRaw);
ASSERT_EQ(home.MachineHomingSeqStep, E_MachineHomingTxState.HX0_REPOS, 'N1/cycle : aucun HX1 par geste joystick'); ASSERT_FALSE(home.M3Locked, 'N1/cycle : aucun verrou homing parasite'); ASSERT_TRUE(home.MachineHomed, 'Reference conservee');
ADVANCE_TIME(10000000); bench(RawPosM1 := raw1, RawPosM2 := raw2);
joy(RawX := bench.Operator.JoyXRaw_ANA1, RawY := bench.Operator.JoyYRaw_ANA2, RawButton := bench.Operator.JoyBtnRaw, Cfg := cfg, NeutralXMem := nx, NeutralYMem := ny);
home(DeadmanArmed := joy.DeadmanArmed, JoystickDeflected := NOT joy.AtNeutralXY, JoystickPull := joy.AxisCmdY.DirectionPositive, JoystickPush := joy.AxisCmdY.DirectionNegative, BtnValidation := bench.Operator.JoyBtnRaw);
ASSERT_EQ(home.MachineHomingSeqStep, E_MachineHomingTxState.HX0_REPOS, 'N1/cycle : aucun HX1 par geste joystick'); ASSERT_FALSE(home.M3Locked, 'N1/cycle : aucun verrou homing parasite'); ASSERT_TRUE(home.MachineHomed, 'Reference conservee');
ADVANCE_TIME(10000000); bench(RawPosM1 := raw1, RawPosM2 := raw2);
joy(RawX := bench.Operator.JoyXRaw_ANA1, RawY := bench.Operator.JoyYRaw_ANA2, RawButton := bench.Operator.JoyBtnRaw, Cfg := cfg, NeutralXMem := nx, NeutralYMem := ny);
home(DeadmanArmed := joy.DeadmanArmed, JoystickDeflected := NOT joy.AtNeutralXY, JoystickPull := joy.AxisCmdY.DirectionPositive, JoystickPush := joy.AxisCmdY.DirectionNegative, BtnValidation := bench.Operator.JoyBtnRaw);
ASSERT_EQ(home.MachineHomingSeqStep, E_MachineHomingTxState.HX0_REPOS, 'N1/cycle : aucun HX1 par geste joystick'); ASSERT_FALSE(home.M3Locked, 'N1/cycle : aucun verrou homing parasite'); ASSERT_TRUE(home.MachineHomed, 'Reference conservee');
ADVANCE_TIME(10000000); bench(RawPosM1 := raw1, RawPosM2 := raw2);
joy(RawX := bench.Operator.JoyXRaw_ANA1, RawY := bench.Operator.JoyYRaw_ANA2, RawButton := bench.Operator.JoyBtnRaw, Cfg := cfg, NeutralXMem := nx, NeutralYMem := ny);
home(DeadmanArmed := joy.DeadmanArmed, JoystickDeflected := NOT joy.AtNeutralXY, JoystickPull := joy.AxisCmdY.DirectionPositive, JoystickPush := joy.AxisCmdY.DirectionNegative, BtnValidation := bench.Operator.JoyBtnRaw);
ASSERT_EQ(home.MachineHomingSeqStep, E_MachineHomingTxState.HX0_REPOS, 'N1/cycle : aucun HX1 par geste joystick'); ASSERT_FALSE(home.M3Locked, 'N1/cycle : aucun verrou homing parasite'); ASSERT_TRUE(home.MachineHomed, 'Reference conservee');
ADVANCE_TIME(10000000); bench(RawPosM1 := raw1, RawPosM2 := raw2);
joy(RawX := bench.Operator.JoyXRaw_ANA1, RawY := bench.Operator.JoyYRaw_ANA2, RawButton := bench.Operator.JoyBtnRaw, Cfg := cfg, NeutralXMem := nx, NeutralYMem := ny);
home(DeadmanArmed := joy.DeadmanArmed, JoystickDeflected := NOT joy.AtNeutralXY, JoystickPull := joy.AxisCmdY.DirectionPositive, JoystickPush := joy.AxisCmdY.DirectionNegative, BtnValidation := bench.Operator.JoyBtnRaw);
ASSERT_EQ(home.MachineHomingSeqStep, E_MachineHomingTxState.HX0_REPOS, 'N1/cycle : aucun HX1 par geste joystick'); ASSERT_FALSE(home.M3Locked, 'N1/cycle : aucun verrou homing parasite'); ASSERT_TRUE(home.MachineHomed, 'Reference conservee');
ADVANCE_TIME(10000000); bench(RawPosM1 := raw1, RawPosM2 := raw2);
joy(RawX := bench.Operator.JoyXRaw_ANA1, RawY := bench.Operator.JoyYRaw_ANA2, RawButton := bench.Operator.JoyBtnRaw, Cfg := cfg, NeutralXMem := nx, NeutralYMem := ny);
home(DeadmanArmed := joy.DeadmanArmed, JoystickDeflected := NOT joy.AtNeutralXY, JoystickPull := joy.AxisCmdY.DirectionPositive, JoystickPush := joy.AxisCmdY.DirectionNegative, BtnValidation := bench.Operator.JoyBtnRaw);
ASSERT_EQ(home.MachineHomingSeqStep, E_MachineHomingTxState.HX0_REPOS, 'N1/cycle : aucun HX1 par geste joystick'); ASSERT_FALSE(home.M3Locked, 'N1/cycle : aucun verrou homing parasite'); ASSERT_TRUE(home.MachineHomed, 'Reference conservee');
ASSERT_TRUE(joy.AxisCmdY.StartStop, 'Geste joystick N1 disponible');
bench.SimJoystickFwd_Up_Close_Active := FALSE;
ADVANCE_TIME(10000000); bench(RawPosM1 := raw1, RawPosM2 := raw2);
joy(RawX := bench.Operator.JoyXRaw_ANA1, RawY := bench.Operator.JoyYRaw_ANA2, RawButton := bench.Operator.JoyBtnRaw, Cfg := cfg, NeutralXMem := nx, NeutralYMem := ny);
home(DeadmanArmed := joy.DeadmanArmed, JoystickDeflected := NOT joy.AtNeutralXY, JoystickPull := joy.AxisCmdY.DirectionPositive, JoystickPush := joy.AxisCmdY.DirectionNegative, BtnValidation := bench.Operator.JoyBtnRaw);
ASSERT_EQ(home.MachineHomingSeqStep, E_MachineHomingTxState.HX0_REPOS, 'N1/cycle : aucun HX1 par geste joystick'); ASSERT_FALSE(home.M3Locked, 'N1/cycle : aucun verrou homing parasite'); ASSERT_TRUE(home.MachineHomed, 'Reference conservee');
ADVANCE_TIME(10000000); bench(RawPosM1 := raw1, RawPosM2 := raw2);
joy(RawX := bench.Operator.JoyXRaw_ANA1, RawY := bench.Operator.JoyYRaw_ANA2, RawButton := bench.Operator.JoyBtnRaw, Cfg := cfg, NeutralXMem := nx, NeutralYMem := ny);
home(DeadmanArmed := joy.DeadmanArmed, JoystickDeflected := NOT joy.AtNeutralXY, JoystickPull := joy.AxisCmdY.DirectionPositive, JoystickPush := joy.AxisCmdY.DirectionNegative, BtnValidation := bench.Operator.JoyBtnRaw);
ASSERT_EQ(home.MachineHomingSeqStep, E_MachineHomingTxState.HX0_REPOS, 'N1/cycle : aucun HX1 par geste joystick'); ASSERT_FALSE(home.M3Locked, 'N1/cycle : aucun verrou homing parasite'); ASSERT_TRUE(home.MachineHomed, 'Reference conservee');
ADVANCE_TIME(10000000); bench(RawPosM1 := raw1, RawPosM2 := raw2);
joy(RawX := bench.Operator.JoyXRaw_ANA1, RawY := bench.Operator.JoyYRaw_ANA2, RawButton := bench.Operator.JoyBtnRaw, Cfg := cfg, NeutralXMem := nx, NeutralYMem := ny);
home(DeadmanArmed := joy.DeadmanArmed, JoystickDeflected := NOT joy.AtNeutralXY, JoystickPull := joy.AxisCmdY.DirectionPositive, JoystickPush := joy.AxisCmdY.DirectionNegative, BtnValidation := bench.Operator.JoyBtnRaw);
ASSERT_EQ(home.MachineHomingSeqStep, E_MachineHomingTxState.HX0_REPOS, 'N1/cycle : aucun HX1 par geste joystick'); ASSERT_FALSE(home.M3Locked, 'N1/cycle : aucun verrou homing parasite'); ASSERT_TRUE(home.MachineHomed, 'Reference conservee');
ADVANCE_TIME(10000000); bench(RawPosM1 := raw1, RawPosM2 := raw2);
joy(RawX := bench.Operator.JoyXRaw_ANA1, RawY := bench.Operator.JoyYRaw_ANA2, RawButton := bench.Operator.JoyBtnRaw, Cfg := cfg, NeutralXMem := nx, NeutralYMem := ny);
home(DeadmanArmed := joy.DeadmanArmed, JoystickDeflected := NOT joy.AtNeutralXY, JoystickPull := joy.AxisCmdY.DirectionPositive, JoystickPush := joy.AxisCmdY.DirectionNegative, BtnValidation := bench.Operator.JoyBtnRaw);
ASSERT_EQ(home.MachineHomingSeqStep, E_MachineHomingTxState.HX0_REPOS, 'N1/cycle : aucun HX1 par geste joystick'); ASSERT_FALSE(home.M3Locked, 'N1/cycle : aucun verrou homing parasite'); ASSERT_TRUE(home.MachineHomed, 'Reference conservee');
ADVANCE_TIME(10000000); bench(RawPosM1 := raw1, RawPosM2 := raw2);
joy(RawX := bench.Operator.JoyXRaw_ANA1, RawY := bench.Operator.JoyYRaw_ANA2, RawButton := bench.Operator.JoyBtnRaw, Cfg := cfg, NeutralXMem := nx, NeutralYMem := ny);
home(DeadmanArmed := joy.DeadmanArmed, JoystickDeflected := NOT joy.AtNeutralXY, JoystickPull := joy.AxisCmdY.DirectionPositive, JoystickPush := joy.AxisCmdY.DirectionNegative, BtnValidation := bench.Operator.JoyBtnRaw);
ASSERT_EQ(home.MachineHomingSeqStep, E_MachineHomingTxState.HX0_REPOS, 'N1/cycle : aucun HX1 par geste joystick'); ASSERT_FALSE(home.M3Locked, 'N1/cycle : aucun verrou homing parasite'); ASSERT_TRUE(home.MachineHomed, 'Reference conservee');
ADVANCE_TIME(10000000); bench(RawPosM1 := raw1, RawPosM2 := raw2);
joy(RawX := bench.Operator.JoyXRaw_ANA1, RawY := bench.Operator.JoyYRaw_ANA2, RawButton := bench.Operator.JoyBtnRaw, Cfg := cfg, NeutralXMem := nx, NeutralYMem := ny);
home(DeadmanArmed := joy.DeadmanArmed, JoystickDeflected := NOT joy.AtNeutralXY, JoystickPull := joy.AxisCmdY.DirectionPositive, JoystickPush := joy.AxisCmdY.DirectionNegative, BtnValidation := bench.Operator.JoyBtnRaw);
ASSERT_EQ(home.MachineHomingSeqStep, E_MachineHomingTxState.HX0_REPOS, 'N1/cycle : aucun HX1 par geste joystick'); ASSERT_FALSE(home.M3Locked, 'N1/cycle : aucun verrou homing parasite'); ASSERT_TRUE(home.MachineHomed, 'Reference conservee');
ADVANCE_TIME(10000000); bench(RawPosM1 := raw1, RawPosM2 := raw2);
joy(RawX := bench.Operator.JoyXRaw_ANA1, RawY := bench.Operator.JoyYRaw_ANA2, RawButton := bench.Operator.JoyBtnRaw, Cfg := cfg, NeutralXMem := nx, NeutralYMem := ny);
home(DeadmanArmed := joy.DeadmanArmed, JoystickDeflected := NOT joy.AtNeutralXY, JoystickPull := joy.AxisCmdY.DirectionPositive, JoystickPush := joy.AxisCmdY.DirectionNegative, BtnValidation := bench.Operator.JoyBtnRaw);
ASSERT_EQ(home.MachineHomingSeqStep, E_MachineHomingTxState.HX0_REPOS, 'N1/cycle : aucun HX1 par geste joystick'); ASSERT_FALSE(home.M3Locked, 'N1/cycle : aucun verrou homing parasite'); ASSERT_TRUE(home.MachineHomed, 'Reference conservee');
ADVANCE_TIME(10000000); bench(RawPosM1 := raw1, RawPosM2 := raw2);
joy(RawX := bench.Operator.JoyXRaw_ANA1, RawY := bench.Operator.JoyYRaw_ANA2, RawButton := bench.Operator.JoyBtnRaw, Cfg := cfg, NeutralXMem := nx, NeutralYMem := ny);
home(DeadmanArmed := joy.DeadmanArmed, JoystickDeflected := NOT joy.AtNeutralXY, JoystickPull := joy.AxisCmdY.DirectionPositive, JoystickPush := joy.AxisCmdY.DirectionNegative, BtnValidation := bench.Operator.JoyBtnRaw);
ASSERT_EQ(home.MachineHomingSeqStep, E_MachineHomingTxState.HX0_REPOS, 'N1/cycle : aucun HX1 par geste joystick'); ASSERT_FALSE(home.M3Locked, 'N1/cycle : aucun verrou homing parasite'); ASSERT_TRUE(home.MachineHomed, 'Reference conservee');
ADVANCE_TIME(10000000); bench(RawPosM1 := raw1, RawPosM2 := raw2);
joy(RawX := bench.Operator.JoyXRaw_ANA1, RawY := bench.Operator.JoyYRaw_ANA2, RawButton := bench.Operator.JoyBtnRaw, Cfg := cfg, NeutralXMem := nx, NeutralYMem := ny);
home(DeadmanArmed := joy.DeadmanArmed, JoystickDeflected := NOT joy.AtNeutralXY, JoystickPull := joy.AxisCmdY.DirectionPositive, JoystickPush := joy.AxisCmdY.DirectionNegative, BtnValidation := bench.Operator.JoyBtnRaw);
ASSERT_EQ(home.MachineHomingSeqStep, E_MachineHomingTxState.HX0_REPOS, 'N1/cycle : aucun HX1 par geste joystick'); ASSERT_FALSE(home.M3Locked, 'N1/cycle : aucun verrou homing parasite'); ASSERT_TRUE(home.MachineHomed, 'Reference conservee');
ADVANCE_TIME(10000000); bench(RawPosM1 := raw1, RawPosM2 := raw2);
joy(RawX := bench.Operator.JoyXRaw_ANA1, RawY := bench.Operator.JoyYRaw_ANA2, RawButton := bench.Operator.JoyBtnRaw, Cfg := cfg, NeutralXMem := nx, NeutralYMem := ny);
home(DeadmanArmed := joy.DeadmanArmed, JoystickDeflected := NOT joy.AtNeutralXY, JoystickPull := joy.AxisCmdY.DirectionPositive, JoystickPush := joy.AxisCmdY.DirectionNegative, BtnValidation := bench.Operator.JoyBtnRaw);
ASSERT_EQ(home.MachineHomingSeqStep, E_MachineHomingTxState.HX0_REPOS, 'N1/cycle : aucun HX1 par geste joystick'); ASSERT_FALSE(home.M3Locked, 'N1/cycle : aucun verrou homing parasite'); ASSERT_TRUE(home.MachineHomed, 'Reference conservee');
ADVANCE_TIME(10000000); bench(RawPosM1 := raw1, RawPosM2 := raw2);
joy(RawX := bench.Operator.JoyXRaw_ANA1, RawY := bench.Operator.JoyYRaw_ANA2, RawButton := bench.Operator.JoyBtnRaw, Cfg := cfg, NeutralXMem := nx, NeutralYMem := ny);
home(DeadmanArmed := joy.DeadmanArmed, JoystickDeflected := NOT joy.AtNeutralXY, JoystickPull := joy.AxisCmdY.DirectionPositive, JoystickPush := joy.AxisCmdY.DirectionNegative, BtnValidation := bench.Operator.JoyBtnRaw);
ASSERT_EQ(home.MachineHomingSeqStep, E_MachineHomingTxState.HX0_REPOS, 'N1/cycle : aucun HX1 par geste joystick'); ASSERT_FALSE(home.M3Locked, 'N1/cycle : aucun verrou homing parasite'); ASSERT_TRUE(home.MachineHomed, 'Reference conservee');
ADVANCE_TIME(10000000); bench(RawPosM1 := raw1, RawPosM2 := raw2);
joy(RawX := bench.Operator.JoyXRaw_ANA1, RawY := bench.Operator.JoyYRaw_ANA2, RawButton := bench.Operator.JoyBtnRaw, Cfg := cfg, NeutralXMem := nx, NeutralYMem := ny);
home(DeadmanArmed := joy.DeadmanArmed, JoystickDeflected := NOT joy.AtNeutralXY, JoystickPull := joy.AxisCmdY.DirectionPositive, JoystickPush := joy.AxisCmdY.DirectionNegative, BtnValidation := bench.Operator.JoyBtnRaw);
ASSERT_EQ(home.MachineHomingSeqStep, E_MachineHomingTxState.HX0_REPOS, 'N1/cycle : aucun HX1 par geste joystick'); ASSERT_FALSE(home.M3Locked, 'N1/cycle : aucun verrou homing parasite'); ASSERT_TRUE(home.MachineHomed, 'Reference conservee');
ADVANCE_TIME(10000000); bench(RawPosM1 := raw1, RawPosM2 := raw2);
joy(RawX := bench.Operator.JoyXRaw_ANA1, RawY := bench.Operator.JoyYRaw_ANA2, RawButton := bench.Operator.JoyBtnRaw, Cfg := cfg, NeutralXMem := nx, NeutralYMem := ny);
home(DeadmanArmed := joy.DeadmanArmed, JoystickDeflected := NOT joy.AtNeutralXY, JoystickPull := joy.AxisCmdY.DirectionPositive, JoystickPush := joy.AxisCmdY.DirectionNegative, BtnValidation := bench.Operator.JoyBtnRaw);
ASSERT_EQ(home.MachineHomingSeqStep, E_MachineHomingTxState.HX0_REPOS, 'N1/cycle : aucun HX1 par geste joystick'); ASSERT_FALSE(home.M3Locked, 'N1/cycle : aucun verrou homing parasite'); ASSERT_TRUE(home.MachineHomed, 'Reference conservee');
ADVANCE_TIME(10000000); bench(RawPosM1 := raw1, RawPosM2 := raw2);
joy(RawX := bench.Operator.JoyXRaw_ANA1, RawY := bench.Operator.JoyYRaw_ANA2, RawButton := bench.Operator.JoyBtnRaw, Cfg := cfg, NeutralXMem := nx, NeutralYMem := ny);
home(DeadmanArmed := joy.DeadmanArmed, JoystickDeflected := NOT joy.AtNeutralXY, JoystickPull := joy.AxisCmdY.DirectionPositive, JoystickPush := joy.AxisCmdY.DirectionNegative, BtnValidation := bench.Operator.JoyBtnRaw);
ASSERT_EQ(home.MachineHomingSeqStep, E_MachineHomingTxState.HX0_REPOS, 'N1/cycle : aucun HX1 par geste joystick'); ASSERT_FALSE(home.M3Locked, 'N1/cycle : aucun verrou homing parasite'); ASSERT_TRUE(home.MachineHomed, 'Reference conservee');
ADVANCE_TIME(10000000); bench(RawPosM1 := raw1, RawPosM2 := raw2);
joy(RawX := bench.Operator.JoyXRaw_ANA1, RawY := bench.Operator.JoyYRaw_ANA2, RawButton := bench.Operator.JoyBtnRaw, Cfg := cfg, NeutralXMem := nx, NeutralYMem := ny);
home(DeadmanArmed := joy.DeadmanArmed, JoystickDeflected := NOT joy.AtNeutralXY, JoystickPull := joy.AxisCmdY.DirectionPositive, JoystickPush := joy.AxisCmdY.DirectionNegative, BtnValidation := bench.Operator.JoyBtnRaw);
ASSERT_EQ(home.MachineHomingSeqStep, E_MachineHomingTxState.HX0_REPOS, 'N1/cycle : aucun HX1 par geste joystick'); ASSERT_FALSE(home.M3Locked, 'N1/cycle : aucun verrou homing parasite'); ASSERT_TRUE(home.MachineHomed, 'Reference conservee');
ADVANCE_TIME(10000000); bench(RawPosM1 := raw1, RawPosM2 := raw2);
joy(RawX := bench.Operator.JoyXRaw_ANA1, RawY := bench.Operator.JoyYRaw_ANA2, RawButton := bench.Operator.JoyBtnRaw, Cfg := cfg, NeutralXMem := nx, NeutralYMem := ny);
home(DeadmanArmed := joy.DeadmanArmed, JoystickDeflected := NOT joy.AtNeutralXY, JoystickPull := joy.AxisCmdY.DirectionPositive, JoystickPush := joy.AxisCmdY.DirectionNegative, BtnValidation := bench.Operator.JoyBtnRaw);
ASSERT_EQ(home.MachineHomingSeqStep, E_MachineHomingTxState.HX0_REPOS, 'N1/cycle : aucun HX1 par geste joystick'); ASSERT_FALSE(home.M3Locked, 'N1/cycle : aucun verrou homing parasite'); ASSERT_TRUE(home.MachineHomed, 'Reference conservee');
ADVANCE_TIME(10000000); bench(RawPosM1 := raw1, RawPosM2 := raw2);
joy(RawX := bench.Operator.JoyXRaw_ANA1, RawY := bench.Operator.JoyYRaw_ANA2, RawButton := bench.Operator.JoyBtnRaw, Cfg := cfg, NeutralXMem := nx, NeutralYMem := ny);
home(DeadmanArmed := joy.DeadmanArmed, JoystickDeflected := NOT joy.AtNeutralXY, JoystickPull := joy.AxisCmdY.DirectionPositive, JoystickPush := joy.AxisCmdY.DirectionNegative, BtnValidation := bench.Operator.JoyBtnRaw);
ASSERT_EQ(home.MachineHomingSeqStep, E_MachineHomingTxState.HX0_REPOS, 'N1/cycle : aucun HX1 par geste joystick'); ASSERT_FALSE(home.M3Locked, 'N1/cycle : aucun verrou homing parasite'); ASSERT_TRUE(home.MachineHomed, 'Reference conservee');
ADVANCE_TIME(10000000); bench(RawPosM1 := raw1, RawPosM2 := raw2);
joy(RawX := bench.Operator.JoyXRaw_ANA1, RawY := bench.Operator.JoyYRaw_ANA2, RawButton := bench.Operator.JoyBtnRaw, Cfg := cfg, NeutralXMem := nx, NeutralYMem := ny);
home(DeadmanArmed := joy.DeadmanArmed, JoystickDeflected := NOT joy.AtNeutralXY, JoystickPull := joy.AxisCmdY.DirectionPositive, JoystickPush := joy.AxisCmdY.DirectionNegative, BtnValidation := bench.Operator.JoyBtnRaw);
ASSERT_EQ(home.MachineHomingSeqStep, E_MachineHomingTxState.HX0_REPOS, 'N1/cycle : aucun HX1 par geste joystick'); ASSERT_FALSE(home.M3Locked, 'N1/cycle : aucun verrou homing parasite'); ASSERT_TRUE(home.MachineHomed, 'Reference conservee');
ADVANCE_TIME(10000000); bench(RawPosM1 := raw1, RawPosM2 := raw2);
joy(RawX := bench.Operator.JoyXRaw_ANA1, RawY := bench.Operator.JoyYRaw_ANA2, RawButton := bench.Operator.JoyBtnRaw, Cfg := cfg, NeutralXMem := nx, NeutralYMem := ny);
home(DeadmanArmed := joy.DeadmanArmed, JoystickDeflected := NOT joy.AtNeutralXY, JoystickPull := joy.AxisCmdY.DirectionPositive, JoystickPush := joy.AxisCmdY.DirectionNegative, BtnValidation := bench.Operator.JoyBtnRaw);
ASSERT_EQ(home.MachineHomingSeqStep, E_MachineHomingTxState.HX0_REPOS, 'N1/cycle : aucun HX1 par geste joystick'); ASSERT_FALSE(home.M3Locked, 'N1/cycle : aucun verrou homing parasite'); ASSERT_TRUE(home.MachineHomed, 'Reference conservee');
ADVANCE_TIME(10000000); bench(RawPosM1 := raw1, RawPosM2 := raw2);
joy(RawX := bench.Operator.JoyXRaw_ANA1, RawY := bench.Operator.JoyYRaw_ANA2, RawButton := bench.Operator.JoyBtnRaw, Cfg := cfg, NeutralXMem := nx, NeutralYMem := ny);
home(DeadmanArmed := joy.DeadmanArmed, JoystickDeflected := NOT joy.AtNeutralXY, JoystickPull := joy.AxisCmdY.DirectionPositive, JoystickPush := joy.AxisCmdY.DirectionNegative, BtnValidation := bench.Operator.JoyBtnRaw);
ASSERT_EQ(home.MachineHomingSeqStep, E_MachineHomingTxState.HX0_REPOS, 'N1/cycle : aucun HX1 par geste joystick'); ASSERT_FALSE(home.M3Locked, 'N1/cycle : aucun verrou homing parasite'); ASSERT_TRUE(home.MachineHomed, 'Reference conservee');
ADVANCE_TIME(10000000); bench(RawPosM1 := raw1, RawPosM2 := raw2);
joy(RawX := bench.Operator.JoyXRaw_ANA1, RawY := bench.Operator.JoyYRaw_ANA2, RawButton := bench.Operator.JoyBtnRaw, Cfg := cfg, NeutralXMem := nx, NeutralYMem := ny);
home(DeadmanArmed := joy.DeadmanArmed, JoystickDeflected := NOT joy.AtNeutralXY, JoystickPull := joy.AxisCmdY.DirectionPositive, JoystickPush := joy.AxisCmdY.DirectionNegative, BtnValidation := bench.Operator.JoyBtnRaw);
ASSERT_EQ(home.MachineHomingSeqStep, E_MachineHomingTxState.HX0_REPOS, 'N1/cycle : aucun HX1 par geste joystick'); ASSERT_FALSE(home.M3Locked, 'N1/cycle : aucun verrou homing parasite'); ASSERT_TRUE(home.MachineHomed, 'Reference conservee');
ADVANCE_TIME(10000000); bench(RawPosM1 := raw1, RawPosM2 := raw2);
joy(RawX := bench.Operator.JoyXRaw_ANA1, RawY := bench.Operator.JoyYRaw_ANA2, RawButton := bench.Operator.JoyBtnRaw, Cfg := cfg, NeutralXMem := nx, NeutralYMem := ny);
home(DeadmanArmed := joy.DeadmanArmed, JoystickDeflected := NOT joy.AtNeutralXY, JoystickPull := joy.AxisCmdY.DirectionPositive, JoystickPush := joy.AxisCmdY.DirectionNegative, BtnValidation := bench.Operator.JoyBtnRaw);
ASSERT_EQ(home.MachineHomingSeqStep, E_MachineHomingTxState.HX0_REPOS, 'N1/cycle : aucun HX1 par geste joystick'); ASSERT_FALSE(home.M3Locked, 'N1/cycle : aucun verrou homing parasite'); ASSERT_TRUE(home.MachineHomed, 'Reference conservee');
ADVANCE_TIME(10000000); bench(RawPosM1 := raw1, RawPosM2 := raw2);
joy(RawX := bench.Operator.JoyXRaw_ANA1, RawY := bench.Operator.JoyYRaw_ANA2, RawButton := bench.Operator.JoyBtnRaw, Cfg := cfg, NeutralXMem := nx, NeutralYMem := ny);
home(DeadmanArmed := joy.DeadmanArmed, JoystickDeflected := NOT joy.AtNeutralXY, JoystickPull := joy.AxisCmdY.DirectionPositive, JoystickPush := joy.AxisCmdY.DirectionNegative, BtnValidation := bench.Operator.JoyBtnRaw);
ASSERT_EQ(home.MachineHomingSeqStep, E_MachineHomingTxState.HX0_REPOS, 'N1/cycle : aucun HX1 par geste joystick'); ASSERT_FALSE(home.M3Locked, 'N1/cycle : aucun verrou homing parasite'); ASSERT_TRUE(home.MachineHomed, 'Reference conservee');
ADVANCE_TIME(10000000); bench(RawPosM1 := raw1, RawPosM2 := raw2);
joy(RawX := bench.Operator.JoyXRaw_ANA1, RawY := bench.Operator.JoyYRaw_ANA2, RawButton := bench.Operator.JoyBtnRaw, Cfg := cfg, NeutralXMem := nx, NeutralYMem := ny);
home(DeadmanArmed := joy.DeadmanArmed, JoystickDeflected := NOT joy.AtNeutralXY, JoystickPull := joy.AxisCmdY.DirectionPositive, JoystickPush := joy.AxisCmdY.DirectionNegative, BtnValidation := bench.Operator.JoyBtnRaw);
ASSERT_EQ(home.MachineHomingSeqStep, E_MachineHomingTxState.HX0_REPOS, 'N1/cycle : aucun HX1 par geste joystick'); ASSERT_FALSE(home.M3Locked, 'N1/cycle : aucun verrou homing parasite'); ASSERT_TRUE(home.MachineHomed, 'Reference conservee');
ADVANCE_TIME(10000000); bench(RawPosM1 := raw1, RawPosM2 := raw2);
joy(RawX := bench.Operator.JoyXRaw_ANA1, RawY := bench.Operator.JoyYRaw_ANA2, RawButton := bench.Operator.JoyBtnRaw, Cfg := cfg, NeutralXMem := nx, NeutralYMem := ny);
home(DeadmanArmed := joy.DeadmanArmed, JoystickDeflected := NOT joy.AtNeutralXY, JoystickPull := joy.AxisCmdY.DirectionPositive, JoystickPush := joy.AxisCmdY.DirectionNegative, BtnValidation := bench.Operator.JoyBtnRaw);
ASSERT_EQ(home.MachineHomingSeqStep, E_MachineHomingTxState.HX0_REPOS, 'N1/cycle : aucun HX1 par geste joystick'); ASSERT_FALSE(home.M3Locked, 'N1/cycle : aucun verrou homing parasite'); ASSERT_TRUE(home.MachineHomed, 'Reference conservee');
home.Mode := E_Mode.SEMI_AUTO; bench.SimJoystickRev_Down_Open_Active := TRUE;
ADVANCE_TIME(10000000); bench(RawPosM1 := raw1, RawPosM2 := raw2);
joy(RawX := bench.Operator.JoyXRaw_ANA1, RawY := bench.Operator.JoyYRaw_ANA2, RawButton := bench.Operator.JoyBtnRaw, Cfg := cfg, NeutralXMem := nx, NeutralYMem := ny);
home(DeadmanArmed := joy.DeadmanArmed, JoystickDeflected := NOT joy.AtNeutralXY, JoystickPull := joy.AxisCmdY.DirectionPositive, JoystickPush := joy.AxisCmdY.DirectionNegative, BtnValidation := bench.Operator.JoyBtnRaw);
ASSERT_EQ(home.MachineHomingSeqStep, E_MachineHomingTxState.HX0_REPOS, 'N1/cycle : aucun HX1 par geste joystick'); ASSERT_FALSE(home.M3Locked, 'N1/cycle : aucun verrou homing parasite'); ASSERT_TRUE(home.MachineHomed, 'Reference conservee');
ADVANCE_TIME(10000000); bench(RawPosM1 := raw1, RawPosM2 := raw2);
joy(RawX := bench.Operator.JoyXRaw_ANA1, RawY := bench.Operator.JoyYRaw_ANA2, RawButton := bench.Operator.JoyBtnRaw, Cfg := cfg, NeutralXMem := nx, NeutralYMem := ny);
home(DeadmanArmed := joy.DeadmanArmed, JoystickDeflected := NOT joy.AtNeutralXY, JoystickPull := joy.AxisCmdY.DirectionPositive, JoystickPush := joy.AxisCmdY.DirectionNegative, BtnValidation := bench.Operator.JoyBtnRaw);
ASSERT_EQ(home.MachineHomingSeqStep, E_MachineHomingTxState.HX0_REPOS, 'N1/cycle : aucun HX1 par geste joystick'); ASSERT_FALSE(home.M3Locked, 'N1/cycle : aucun verrou homing parasite'); ASSERT_TRUE(home.MachineHomed, 'Reference conservee');
ADVANCE_TIME(10000000); bench(RawPosM1 := raw1, RawPosM2 := raw2);
joy(RawX := bench.Operator.JoyXRaw_ANA1, RawY := bench.Operator.JoyYRaw_ANA2, RawButton := bench.Operator.JoyBtnRaw, Cfg := cfg, NeutralXMem := nx, NeutralYMem := ny);
home(DeadmanArmed := joy.DeadmanArmed, JoystickDeflected := NOT joy.AtNeutralXY, JoystickPull := joy.AxisCmdY.DirectionPositive, JoystickPush := joy.AxisCmdY.DirectionNegative, BtnValidation := bench.Operator.JoyBtnRaw);
ASSERT_EQ(home.MachineHomingSeqStep, E_MachineHomingTxState.HX0_REPOS, 'N1/cycle : aucun HX1 par geste joystick'); ASSERT_FALSE(home.M3Locked, 'N1/cycle : aucun verrou homing parasite'); ASSERT_TRUE(home.MachineHomed, 'Reference conservee');
ADVANCE_TIME(10000000); bench(RawPosM1 := raw1, RawPosM2 := raw2);
joy(RawX := bench.Operator.JoyXRaw_ANA1, RawY := bench.Operator.JoyYRaw_ANA2, RawButton := bench.Operator.JoyBtnRaw, Cfg := cfg, NeutralXMem := nx, NeutralYMem := ny);
home(DeadmanArmed := joy.DeadmanArmed, JoystickDeflected := NOT joy.AtNeutralXY, JoystickPull := joy.AxisCmdY.DirectionPositive, JoystickPush := joy.AxisCmdY.DirectionNegative, BtnValidation := bench.Operator.JoyBtnRaw);
ASSERT_EQ(home.MachineHomingSeqStep, E_MachineHomingTxState.HX0_REPOS, 'N1/cycle : aucun HX1 par geste joystick'); ASSERT_FALSE(home.M3Locked, 'N1/cycle : aucun verrou homing parasite'); ASSERT_TRUE(home.MachineHomed, 'Reference conservee');
ADVANCE_TIME(10000000); bench(RawPosM1 := raw1, RawPosM2 := raw2);
joy(RawX := bench.Operator.JoyXRaw_ANA1, RawY := bench.Operator.JoyYRaw_ANA2, RawButton := bench.Operator.JoyBtnRaw, Cfg := cfg, NeutralXMem := nx, NeutralYMem := ny);
home(DeadmanArmed := joy.DeadmanArmed, JoystickDeflected := NOT joy.AtNeutralXY, JoystickPull := joy.AxisCmdY.DirectionPositive, JoystickPush := joy.AxisCmdY.DirectionNegative, BtnValidation := bench.Operator.JoyBtnRaw);
ASSERT_EQ(home.MachineHomingSeqStep, E_MachineHomingTxState.HX0_REPOS, 'N1/cycle : aucun HX1 par geste joystick'); ASSERT_FALSE(home.M3Locked, 'N1/cycle : aucun verrou homing parasite'); ASSERT_TRUE(home.MachineHomed, 'Reference conservee');
ADVANCE_TIME(10000000); bench(RawPosM1 := raw1, RawPosM2 := raw2);
joy(RawX := bench.Operator.JoyXRaw_ANA1, RawY := bench.Operator.JoyYRaw_ANA2, RawButton := bench.Operator.JoyBtnRaw, Cfg := cfg, NeutralXMem := nx, NeutralYMem := ny);
home(DeadmanArmed := joy.DeadmanArmed, JoystickDeflected := NOT joy.AtNeutralXY, JoystickPull := joy.AxisCmdY.DirectionPositive, JoystickPush := joy.AxisCmdY.DirectionNegative, BtnValidation := bench.Operator.JoyBtnRaw);
ASSERT_EQ(home.MachineHomingSeqStep, E_MachineHomingTxState.HX0_REPOS, 'N1/cycle : aucun HX1 par geste joystick'); ASSERT_FALSE(home.M3Locked, 'N1/cycle : aucun verrou homing parasite'); ASSERT_TRUE(home.MachineHomed, 'Reference conservee');
ADVANCE_TIME(10000000); bench(RawPosM1 := raw1, RawPosM2 := raw2);
joy(RawX := bench.Operator.JoyXRaw_ANA1, RawY := bench.Operator.JoyYRaw_ANA2, RawButton := bench.Operator.JoyBtnRaw, Cfg := cfg, NeutralXMem := nx, NeutralYMem := ny);
home(DeadmanArmed := joy.DeadmanArmed, JoystickDeflected := NOT joy.AtNeutralXY, JoystickPull := joy.AxisCmdY.DirectionPositive, JoystickPush := joy.AxisCmdY.DirectionNegative, BtnValidation := bench.Operator.JoyBtnRaw);
ASSERT_EQ(home.MachineHomingSeqStep, E_MachineHomingTxState.HX0_REPOS, 'N1/cycle : aucun HX1 par geste joystick'); ASSERT_FALSE(home.M3Locked, 'N1/cycle : aucun verrou homing parasite'); ASSERT_TRUE(home.MachineHomed, 'Reference conservee');
ADVANCE_TIME(10000000); bench(RawPosM1 := raw1, RawPosM2 := raw2);
joy(RawX := bench.Operator.JoyXRaw_ANA1, RawY := bench.Operator.JoyYRaw_ANA2, RawButton := bench.Operator.JoyBtnRaw, Cfg := cfg, NeutralXMem := nx, NeutralYMem := ny);
home(DeadmanArmed := joy.DeadmanArmed, JoystickDeflected := NOT joy.AtNeutralXY, JoystickPull := joy.AxisCmdY.DirectionPositive, JoystickPush := joy.AxisCmdY.DirectionNegative, BtnValidation := bench.Operator.JoyBtnRaw);
ASSERT_EQ(home.MachineHomingSeqStep, E_MachineHomingTxState.HX0_REPOS, 'N1/cycle : aucun HX1 par geste joystick'); ASSERT_FALSE(home.M3Locked, 'N1/cycle : aucun verrou homing parasite'); ASSERT_TRUE(home.MachineHomed, 'Reference conservee');
ADVANCE_TIME(10000000); bench(RawPosM1 := raw1, RawPosM2 := raw2);
joy(RawX := bench.Operator.JoyXRaw_ANA1, RawY := bench.Operator.JoyYRaw_ANA2, RawButton := bench.Operator.JoyBtnRaw, Cfg := cfg, NeutralXMem := nx, NeutralYMem := ny);
home(DeadmanArmed := joy.DeadmanArmed, JoystickDeflected := NOT joy.AtNeutralXY, JoystickPull := joy.AxisCmdY.DirectionPositive, JoystickPush := joy.AxisCmdY.DirectionNegative, BtnValidation := bench.Operator.JoyBtnRaw);
ASSERT_EQ(home.MachineHomingSeqStep, E_MachineHomingTxState.HX0_REPOS, 'N1/cycle : aucun HX1 par geste joystick'); ASSERT_FALSE(home.M3Locked, 'N1/cycle : aucun verrou homing parasite'); ASSERT_TRUE(home.MachineHomed, 'Reference conservee');
ADVANCE_TIME(10000000); bench(RawPosM1 := raw1, RawPosM2 := raw2);
joy(RawX := bench.Operator.JoyXRaw_ANA1, RawY := bench.Operator.JoyYRaw_ANA2, RawButton := bench.Operator.JoyBtnRaw, Cfg := cfg, NeutralXMem := nx, NeutralYMem := ny);
home(DeadmanArmed := joy.DeadmanArmed, JoystickDeflected := NOT joy.AtNeutralXY, JoystickPull := joy.AxisCmdY.DirectionPositive, JoystickPush := joy.AxisCmdY.DirectionNegative, BtnValidation := bench.Operator.JoyBtnRaw);
ASSERT_EQ(home.MachineHomingSeqStep, E_MachineHomingTxState.HX0_REPOS, 'N1/cycle : aucun HX1 par geste joystick'); ASSERT_FALSE(home.M3Locked, 'N1/cycle : aucun verrou homing parasite'); ASSERT_TRUE(home.MachineHomed, 'Reference conservee');
ADVANCE_TIME(10000000); bench(RawPosM1 := raw1, RawPosM2 := raw2);
joy(RawX := bench.Operator.JoyXRaw_ANA1, RawY := bench.Operator.JoyYRaw_ANA2, RawButton := bench.Operator.JoyBtnRaw, Cfg := cfg, NeutralXMem := nx, NeutralYMem := ny);
home(DeadmanArmed := joy.DeadmanArmed, JoystickDeflected := NOT joy.AtNeutralXY, JoystickPull := joy.AxisCmdY.DirectionPositive, JoystickPush := joy.AxisCmdY.DirectionNegative, BtnValidation := bench.Operator.JoyBtnRaw);
ASSERT_EQ(home.MachineHomingSeqStep, E_MachineHomingTxState.HX0_REPOS, 'N1/cycle : aucun HX1 par geste joystick'); ASSERT_FALSE(home.M3Locked, 'N1/cycle : aucun verrou homing parasite'); ASSERT_TRUE(home.MachineHomed, 'Reference conservee');
ADVANCE_TIME(10000000); bench(RawPosM1 := raw1, RawPosM2 := raw2);
joy(RawX := bench.Operator.JoyXRaw_ANA1, RawY := bench.Operator.JoyYRaw_ANA2, RawButton := bench.Operator.JoyBtnRaw, Cfg := cfg, NeutralXMem := nx, NeutralYMem := ny);
home(DeadmanArmed := joy.DeadmanArmed, JoystickDeflected := NOT joy.AtNeutralXY, JoystickPull := joy.AxisCmdY.DirectionPositive, JoystickPush := joy.AxisCmdY.DirectionNegative, BtnValidation := bench.Operator.JoyBtnRaw);
ASSERT_EQ(home.MachineHomingSeqStep, E_MachineHomingTxState.HX0_REPOS, 'N1/cycle : aucun HX1 par geste joystick'); ASSERT_FALSE(home.M3Locked, 'N1/cycle : aucun verrou homing parasite'); ASSERT_TRUE(home.MachineHomed, 'Reference conservee');
ADVANCE_TIME(10000000); bench(RawPosM1 := raw1, RawPosM2 := raw2);
joy(RawX := bench.Operator.JoyXRaw_ANA1, RawY := bench.Operator.JoyYRaw_ANA2, RawButton := bench.Operator.JoyBtnRaw, Cfg := cfg, NeutralXMem := nx, NeutralYMem := ny);
home(DeadmanArmed := joy.DeadmanArmed, JoystickDeflected := NOT joy.AtNeutralXY, JoystickPull := joy.AxisCmdY.DirectionPositive, JoystickPush := joy.AxisCmdY.DirectionNegative, BtnValidation := bench.Operator.JoyBtnRaw);
ASSERT_EQ(home.MachineHomingSeqStep, E_MachineHomingTxState.HX0_REPOS, 'N1/cycle : aucun HX1 par geste joystick'); ASSERT_FALSE(home.M3Locked, 'N1/cycle : aucun verrou homing parasite'); ASSERT_TRUE(home.MachineHomed, 'Reference conservee');
ADVANCE_TIME(10000000); bench(RawPosM1 := raw1, RawPosM2 := raw2);
joy(RawX := bench.Operator.JoyXRaw_ANA1, RawY := bench.Operator.JoyYRaw_ANA2, RawButton := bench.Operator.JoyBtnRaw, Cfg := cfg, NeutralXMem := nx, NeutralYMem := ny);
home(DeadmanArmed := joy.DeadmanArmed, JoystickDeflected := NOT joy.AtNeutralXY, JoystickPull := joy.AxisCmdY.DirectionPositive, JoystickPush := joy.AxisCmdY.DirectionNegative, BtnValidation := bench.Operator.JoyBtnRaw);
ASSERT_EQ(home.MachineHomingSeqStep, E_MachineHomingTxState.HX0_REPOS, 'N1/cycle : aucun HX1 par geste joystick'); ASSERT_FALSE(home.M3Locked, 'N1/cycle : aucun verrou homing parasite'); ASSERT_TRUE(home.MachineHomed, 'Reference conservee');
ADVANCE_TIME(10000000); bench(RawPosM1 := raw1, RawPosM2 := raw2);
joy(RawX := bench.Operator.JoyXRaw_ANA1, RawY := bench.Operator.JoyYRaw_ANA2, RawButton := bench.Operator.JoyBtnRaw, Cfg := cfg, NeutralXMem := nx, NeutralYMem := ny);
home(DeadmanArmed := joy.DeadmanArmed, JoystickDeflected := NOT joy.AtNeutralXY, JoystickPull := joy.AxisCmdY.DirectionPositive, JoystickPush := joy.AxisCmdY.DirectionNegative, BtnValidation := bench.Operator.JoyBtnRaw);
ASSERT_EQ(home.MachineHomingSeqStep, E_MachineHomingTxState.HX0_REPOS, 'N1/cycle : aucun HX1 par geste joystick'); ASSERT_FALSE(home.M3Locked, 'N1/cycle : aucun verrou homing parasite'); ASSERT_TRUE(home.MachineHomed, 'Reference conservee');
ADVANCE_TIME(10000000); bench(RawPosM1 := raw1, RawPosM2 := raw2);
joy(RawX := bench.Operator.JoyXRaw_ANA1, RawY := bench.Operator.JoyYRaw_ANA2, RawButton := bench.Operator.JoyBtnRaw, Cfg := cfg, NeutralXMem := nx, NeutralYMem := ny);
home(DeadmanArmed := joy.DeadmanArmed, JoystickDeflected := NOT joy.AtNeutralXY, JoystickPull := joy.AxisCmdY.DirectionPositive, JoystickPush := joy.AxisCmdY.DirectionNegative, BtnValidation := bench.Operator.JoyBtnRaw);
ASSERT_EQ(home.MachineHomingSeqStep, E_MachineHomingTxState.HX0_REPOS, 'N1/cycle : aucun HX1 par geste joystick'); ASSERT_FALSE(home.M3Locked, 'N1/cycle : aucun verrou homing parasite'); ASSERT_TRUE(home.MachineHomed, 'Reference conservee');
ADVANCE_TIME(10000000); bench(RawPosM1 := raw1, RawPosM2 := raw2);
joy(RawX := bench.Operator.JoyXRaw_ANA1, RawY := bench.Operator.JoyYRaw_ANA2, RawButton := bench.Operator.JoyBtnRaw, Cfg := cfg, NeutralXMem := nx, NeutralYMem := ny);
home(DeadmanArmed := joy.DeadmanArmed, JoystickDeflected := NOT joy.AtNeutralXY, JoystickPull := joy.AxisCmdY.DirectionPositive, JoystickPush := joy.AxisCmdY.DirectionNegative, BtnValidation := bench.Operator.JoyBtnRaw);
ASSERT_EQ(home.MachineHomingSeqStep, E_MachineHomingTxState.HX0_REPOS, 'N1/cycle : aucun HX1 par geste joystick'); ASSERT_FALSE(home.M3Locked, 'N1/cycle : aucun verrou homing parasite'); ASSERT_TRUE(home.MachineHomed, 'Reference conservee');
ADVANCE_TIME(10000000); bench(RawPosM1 := raw1, RawPosM2 := raw2);
joy(RawX := bench.Operator.JoyXRaw_ANA1, RawY := bench.Operator.JoyYRaw_ANA2, RawButton := bench.Operator.JoyBtnRaw, Cfg := cfg, NeutralXMem := nx, NeutralYMem := ny);
home(DeadmanArmed := joy.DeadmanArmed, JoystickDeflected := NOT joy.AtNeutralXY, JoystickPull := joy.AxisCmdY.DirectionPositive, JoystickPush := joy.AxisCmdY.DirectionNegative, BtnValidation := bench.Operator.JoyBtnRaw);
ASSERT_EQ(home.MachineHomingSeqStep, E_MachineHomingTxState.HX0_REPOS, 'N1/cycle : aucun HX1 par geste joystick'); ASSERT_FALSE(home.M3Locked, 'N1/cycle : aucun verrou homing parasite'); ASSERT_TRUE(home.MachineHomed, 'Reference conservee');
ADVANCE_TIME(10000000); bench(RawPosM1 := raw1, RawPosM2 := raw2);
joy(RawX := bench.Operator.JoyXRaw_ANA1, RawY := bench.Operator.JoyYRaw_ANA2, RawButton := bench.Operator.JoyBtnRaw, Cfg := cfg, NeutralXMem := nx, NeutralYMem := ny);
home(DeadmanArmed := joy.DeadmanArmed, JoystickDeflected := NOT joy.AtNeutralXY, JoystickPull := joy.AxisCmdY.DirectionPositive, JoystickPush := joy.AxisCmdY.DirectionNegative, BtnValidation := bench.Operator.JoyBtnRaw);
ASSERT_EQ(home.MachineHomingSeqStep, E_MachineHomingTxState.HX0_REPOS, 'N1/cycle : aucun HX1 par geste joystick'); ASSERT_FALSE(home.M3Locked, 'N1/cycle : aucun verrou homing parasite'); ASSERT_TRUE(home.MachineHomed, 'Reference conservee');
ADVANCE_TIME(10000000); bench(RawPosM1 := raw1, RawPosM2 := raw2);
joy(RawX := bench.Operator.JoyXRaw_ANA1, RawY := bench.Operator.JoyYRaw_ANA2, RawButton := bench.Operator.JoyBtnRaw, Cfg := cfg, NeutralXMem := nx, NeutralYMem := ny);
home(DeadmanArmed := joy.DeadmanArmed, JoystickDeflected := NOT joy.AtNeutralXY, JoystickPull := joy.AxisCmdY.DirectionPositive, JoystickPush := joy.AxisCmdY.DirectionNegative, BtnValidation := bench.Operator.JoyBtnRaw);
ASSERT_EQ(home.MachineHomingSeqStep, E_MachineHomingTxState.HX0_REPOS, 'N1/cycle : aucun HX1 par geste joystick'); ASSERT_FALSE(home.M3Locked, 'N1/cycle : aucun verrou homing parasite'); ASSERT_TRUE(home.MachineHomed, 'Reference conservee');
ADVANCE_TIME(10000000); bench(RawPosM1 := raw1, RawPosM2 := raw2);
joy(RawX := bench.Operator.JoyXRaw_ANA1, RawY := bench.Operator.JoyYRaw_ANA2, RawButton := bench.Operator.JoyBtnRaw, Cfg := cfg, NeutralXMem := nx, NeutralYMem := ny);
home(DeadmanArmed := joy.DeadmanArmed, JoystickDeflected := NOT joy.AtNeutralXY, JoystickPull := joy.AxisCmdY.DirectionPositive, JoystickPush := joy.AxisCmdY.DirectionNegative, BtnValidation := bench.Operator.JoyBtnRaw);
ASSERT_EQ(home.MachineHomingSeqStep, E_MachineHomingTxState.HX0_REPOS, 'N1/cycle : aucun HX1 par geste joystick'); ASSERT_FALSE(home.M3Locked, 'N1/cycle : aucun verrou homing parasite'); ASSERT_TRUE(home.MachineHomed, 'Reference conservee');
ADVANCE_TIME(10000000); bench(RawPosM1 := raw1, RawPosM2 := raw2);
joy(RawX := bench.Operator.JoyXRaw_ANA1, RawY := bench.Operator.JoyYRaw_ANA2, RawButton := bench.Operator.JoyBtnRaw, Cfg := cfg, NeutralXMem := nx, NeutralYMem := ny);
home(DeadmanArmed := joy.DeadmanArmed, JoystickDeflected := NOT joy.AtNeutralXY, JoystickPull := joy.AxisCmdY.DirectionPositive, JoystickPush := joy.AxisCmdY.DirectionNegative, BtnValidation := bench.Operator.JoyBtnRaw);
ASSERT_EQ(home.MachineHomingSeqStep, E_MachineHomingTxState.HX0_REPOS, 'N1/cycle : aucun HX1 par geste joystick'); ASSERT_FALSE(home.M3Locked, 'N1/cycle : aucun verrou homing parasite'); ASSERT_TRUE(home.MachineHomed, 'Reference conservee');
ADVANCE_TIME(10000000); bench(RawPosM1 := raw1, RawPosM2 := raw2);
joy(RawX := bench.Operator.JoyXRaw_ANA1, RawY := bench.Operator.JoyYRaw_ANA2, RawButton := bench.Operator.JoyBtnRaw, Cfg := cfg, NeutralXMem := nx, NeutralYMem := ny);
home(DeadmanArmed := joy.DeadmanArmed, JoystickDeflected := NOT joy.AtNeutralXY, JoystickPull := joy.AxisCmdY.DirectionPositive, JoystickPush := joy.AxisCmdY.DirectionNegative, BtnValidation := bench.Operator.JoyBtnRaw);
ASSERT_EQ(home.MachineHomingSeqStep, E_MachineHomingTxState.HX0_REPOS, 'N1/cycle : aucun HX1 par geste joystick'); ASSERT_FALSE(home.M3Locked, 'N1/cycle : aucun verrou homing parasite'); ASSERT_TRUE(home.MachineHomed, 'Reference conservee');
ADVANCE_TIME(10000000); bench(RawPosM1 := raw1, RawPosM2 := raw2);
joy(RawX := bench.Operator.JoyXRaw_ANA1, RawY := bench.Operator.JoyYRaw_ANA2, RawButton := bench.Operator.JoyBtnRaw, Cfg := cfg, NeutralXMem := nx, NeutralYMem := ny);
home(DeadmanArmed := joy.DeadmanArmed, JoystickDeflected := NOT joy.AtNeutralXY, JoystickPull := joy.AxisCmdY.DirectionPositive, JoystickPush := joy.AxisCmdY.DirectionNegative, BtnValidation := bench.Operator.JoyBtnRaw);
ASSERT_EQ(home.MachineHomingSeqStep, E_MachineHomingTxState.HX0_REPOS, 'N1/cycle : aucun HX1 par geste joystick'); ASSERT_FALSE(home.M3Locked, 'N1/cycle : aucun verrou homing parasite'); ASSERT_TRUE(home.MachineHomed, 'Reference conservee');
ADVANCE_TIME(10000000); bench(RawPosM1 := raw1, RawPosM2 := raw2);
joy(RawX := bench.Operator.JoyXRaw_ANA1, RawY := bench.Operator.JoyYRaw_ANA2, RawButton := bench.Operator.JoyBtnRaw, Cfg := cfg, NeutralXMem := nx, NeutralYMem := ny);
home(DeadmanArmed := joy.DeadmanArmed, JoystickDeflected := NOT joy.AtNeutralXY, JoystickPull := joy.AxisCmdY.DirectionPositive, JoystickPush := joy.AxisCmdY.DirectionNegative, BtnValidation := bench.Operator.JoyBtnRaw);
ASSERT_EQ(home.MachineHomingSeqStep, E_MachineHomingTxState.HX0_REPOS, 'N1/cycle : aucun HX1 par geste joystick'); ASSERT_FALSE(home.M3Locked, 'N1/cycle : aucun verrou homing parasite'); ASSERT_TRUE(home.MachineHomed, 'Reference conservee');
ADVANCE_TIME(10000000); bench(RawPosM1 := raw1, RawPosM2 := raw2);
joy(RawX := bench.Operator.JoyXRaw_ANA1, RawY := bench.Operator.JoyYRaw_ANA2, RawButton := bench.Operator.JoyBtnRaw, Cfg := cfg, NeutralXMem := nx, NeutralYMem := ny);
home(DeadmanArmed := joy.DeadmanArmed, JoystickDeflected := NOT joy.AtNeutralXY, JoystickPull := joy.AxisCmdY.DirectionPositive, JoystickPush := joy.AxisCmdY.DirectionNegative, BtnValidation := bench.Operator.JoyBtnRaw);
ASSERT_EQ(home.MachineHomingSeqStep, E_MachineHomingTxState.HX0_REPOS, 'N1/cycle : aucun HX1 par geste joystick'); ASSERT_FALSE(home.M3Locked, 'N1/cycle : aucun verrou homing parasite'); ASSERT_TRUE(home.MachineHomed, 'Reference conservee');
ADVANCE_TIME(10000000); bench(RawPosM1 := raw1, RawPosM2 := raw2);
joy(RawX := bench.Operator.JoyXRaw_ANA1, RawY := bench.Operator.JoyYRaw_ANA2, RawButton := bench.Operator.JoyBtnRaw, Cfg := cfg, NeutralXMem := nx, NeutralYMem := ny);
home(DeadmanArmed := joy.DeadmanArmed, JoystickDeflected := NOT joy.AtNeutralXY, JoystickPull := joy.AxisCmdY.DirectionPositive, JoystickPush := joy.AxisCmdY.DirectionNegative, BtnValidation := bench.Operator.JoyBtnRaw);
ASSERT_EQ(home.MachineHomingSeqStep, E_MachineHomingTxState.HX0_REPOS, 'N1/cycle : aucun HX1 par geste joystick'); ASSERT_FALSE(home.M3Locked, 'N1/cycle : aucun verrou homing parasite'); ASSERT_TRUE(home.MachineHomed, 'Reference conservee');
ADVANCE_TIME(10000000); bench(RawPosM1 := raw1, RawPosM2 := raw2);
joy(RawX := bench.Operator.JoyXRaw_ANA1, RawY := bench.Operator.JoyYRaw_ANA2, RawButton := bench.Operator.JoyBtnRaw, Cfg := cfg, NeutralXMem := nx, NeutralYMem := ny);
home(DeadmanArmed := joy.DeadmanArmed, JoystickDeflected := NOT joy.AtNeutralXY, JoystickPull := joy.AxisCmdY.DirectionPositive, JoystickPush := joy.AxisCmdY.DirectionNegative, BtnValidation := bench.Operator.JoyBtnRaw);
ASSERT_EQ(home.MachineHomingSeqStep, E_MachineHomingTxState.HX0_REPOS, 'N1/cycle : aucun HX1 par geste joystick'); ASSERT_FALSE(home.M3Locked, 'N1/cycle : aucun verrou homing parasite'); ASSERT_TRUE(home.MachineHomed, 'Reference conservee');
ADVANCE_TIME(10000000); bench(RawPosM1 := raw1, RawPosM2 := raw2);
joy(RawX := bench.Operator.JoyXRaw_ANA1, RawY := bench.Operator.JoyYRaw_ANA2, RawButton := bench.Operator.JoyBtnRaw, Cfg := cfg, NeutralXMem := nx, NeutralYMem := ny);
home(DeadmanArmed := joy.DeadmanArmed, JoystickDeflected := NOT joy.AtNeutralXY, JoystickPull := joy.AxisCmdY.DirectionPositive, JoystickPush := joy.AxisCmdY.DirectionNegative, BtnValidation := bench.Operator.JoyBtnRaw);
ASSERT_EQ(home.MachineHomingSeqStep, E_MachineHomingTxState.HX0_REPOS, 'N1/cycle : aucun HX1 par geste joystick'); ASSERT_FALSE(home.M3Locked, 'N1/cycle : aucun verrou homing parasite'); ASSERT_TRUE(home.MachineHomed, 'Reference conservee');
ADVANCE_TIME(10000000); bench(RawPosM1 := raw1, RawPosM2 := raw2);
joy(RawX := bench.Operator.JoyXRaw_ANA1, RawY := bench.Operator.JoyYRaw_ANA2, RawButton := bench.Operator.JoyBtnRaw, Cfg := cfg, NeutralXMem := nx, NeutralYMem := ny);
home(DeadmanArmed := joy.DeadmanArmed, JoystickDeflected := NOT joy.AtNeutralXY, JoystickPull := joy.AxisCmdY.DirectionPositive, JoystickPush := joy.AxisCmdY.DirectionNegative, BtnValidation := bench.Operator.JoyBtnRaw);
ASSERT_EQ(home.MachineHomingSeqStep, E_MachineHomingTxState.HX0_REPOS, 'N1/cycle : aucun HX1 par geste joystick'); ASSERT_FALSE(home.M3Locked, 'N1/cycle : aucun verrou homing parasite'); ASSERT_TRUE(home.MachineHomed, 'Reference conservee');
ADVANCE_TIME(10000000); bench(RawPosM1 := raw1, RawPosM2 := raw2);
joy(RawX := bench.Operator.JoyXRaw_ANA1, RawY := bench.Operator.JoyYRaw_ANA2, RawButton := bench.Operator.JoyBtnRaw, Cfg := cfg, NeutralXMem := nx, NeutralYMem := ny);
home(DeadmanArmed := joy.DeadmanArmed, JoystickDeflected := NOT joy.AtNeutralXY, JoystickPull := joy.AxisCmdY.DirectionPositive, JoystickPush := joy.AxisCmdY.DirectionNegative, BtnValidation := bench.Operator.JoyBtnRaw);
ASSERT_EQ(home.MachineHomingSeqStep, E_MachineHomingTxState.HX0_REPOS, 'N1/cycle : aucun HX1 par geste joystick'); ASSERT_FALSE(home.M3Locked, 'N1/cycle : aucun verrou homing parasite'); ASSERT_TRUE(home.MachineHomed, 'Reference conservee');
ADVANCE_TIME(10000000); bench(RawPosM1 := raw1, RawPosM2 := raw2);
joy(RawX := bench.Operator.JoyXRaw_ANA1, RawY := bench.Operator.JoyYRaw_ANA2, RawButton := bench.Operator.JoyBtnRaw, Cfg := cfg, NeutralXMem := nx, NeutralYMem := ny);
home(DeadmanArmed := joy.DeadmanArmed, JoystickDeflected := NOT joy.AtNeutralXY, JoystickPull := joy.AxisCmdY.DirectionPositive, JoystickPush := joy.AxisCmdY.DirectionNegative, BtnValidation := bench.Operator.JoyBtnRaw);
ASSERT_EQ(home.MachineHomingSeqStep, E_MachineHomingTxState.HX0_REPOS, 'N1/cycle : aucun HX1 par geste joystick'); ASSERT_FALSE(home.M3Locked, 'N1/cycle : aucun verrou homing parasite'); ASSERT_TRUE(home.MachineHomed, 'Reference conservee');
ADVANCE_TIME(10000000); bench(RawPosM1 := raw1, RawPosM2 := raw2);
joy(RawX := bench.Operator.JoyXRaw_ANA1, RawY := bench.Operator.JoyYRaw_ANA2, RawButton := bench.Operator.JoyBtnRaw, Cfg := cfg, NeutralXMem := nx, NeutralYMem := ny);
home(DeadmanArmed := joy.DeadmanArmed, JoystickDeflected := NOT joy.AtNeutralXY, JoystickPull := joy.AxisCmdY.DirectionPositive, JoystickPush := joy.AxisCmdY.DirectionNegative, BtnValidation := bench.Operator.JoyBtnRaw);
ASSERT_EQ(home.MachineHomingSeqStep, E_MachineHomingTxState.HX0_REPOS, 'N1/cycle : aucun HX1 par geste joystick'); ASSERT_FALSE(home.M3Locked, 'N1/cycle : aucun verrou homing parasite'); ASSERT_TRUE(home.MachineHomed, 'Reference conservee');
ADVANCE_TIME(10000000); bench(RawPosM1 := raw1, RawPosM2 := raw2);
joy(RawX := bench.Operator.JoyXRaw_ANA1, RawY := bench.Operator.JoyYRaw_ANA2, RawButton := bench.Operator.JoyBtnRaw, Cfg := cfg, NeutralXMem := nx, NeutralYMem := ny);
home(DeadmanArmed := joy.DeadmanArmed, JoystickDeflected := NOT joy.AtNeutralXY, JoystickPull := joy.AxisCmdY.DirectionPositive, JoystickPush := joy.AxisCmdY.DirectionNegative, BtnValidation := bench.Operator.JoyBtnRaw);
ASSERT_EQ(home.MachineHomingSeqStep, E_MachineHomingTxState.HX0_REPOS, 'N1/cycle : aucun HX1 par geste joystick'); ASSERT_FALSE(home.M3Locked, 'N1/cycle : aucun verrou homing parasite'); ASSERT_TRUE(home.MachineHomed, 'Reference conservee');
ADVANCE_TIME(10000000); bench(RawPosM1 := raw1, RawPosM2 := raw2);
joy(RawX := bench.Operator.JoyXRaw_ANA1, RawY := bench.Operator.JoyYRaw_ANA2, RawButton := bench.Operator.JoyBtnRaw, Cfg := cfg, NeutralXMem := nx, NeutralYMem := ny);
home(DeadmanArmed := joy.DeadmanArmed, JoystickDeflected := NOT joy.AtNeutralXY, JoystickPull := joy.AxisCmdY.DirectionPositive, JoystickPush := joy.AxisCmdY.DirectionNegative, BtnValidation := bench.Operator.JoyBtnRaw);
ASSERT_EQ(home.MachineHomingSeqStep, E_MachineHomingTxState.HX0_REPOS, 'N1/cycle : aucun HX1 par geste joystick'); ASSERT_FALSE(home.M3Locked, 'N1/cycle : aucun verrou homing parasite'); ASSERT_TRUE(home.MachineHomed, 'Reference conservee');
ADVANCE_TIME(10000000); bench(RawPosM1 := raw1, RawPosM2 := raw2);
joy(RawX := bench.Operator.JoyXRaw_ANA1, RawY := bench.Operator.JoyYRaw_ANA2, RawButton := bench.Operator.JoyBtnRaw, Cfg := cfg, NeutralXMem := nx, NeutralYMem := ny);
home(DeadmanArmed := joy.DeadmanArmed, JoystickDeflected := NOT joy.AtNeutralXY, JoystickPull := joy.AxisCmdY.DirectionPositive, JoystickPush := joy.AxisCmdY.DirectionNegative, BtnValidation := bench.Operator.JoyBtnRaw);
ASSERT_EQ(home.MachineHomingSeqStep, E_MachineHomingTxState.HX0_REPOS, 'N1/cycle : aucun HX1 par geste joystick'); ASSERT_FALSE(home.M3Locked, 'N1/cycle : aucun verrou homing parasite'); ASSERT_TRUE(home.MachineHomed, 'Reference conservee');
ADVANCE_TIME(10000000); bench(RawPosM1 := raw1, RawPosM2 := raw2);
joy(RawX := bench.Operator.JoyXRaw_ANA1, RawY := bench.Operator.JoyYRaw_ANA2, RawButton := bench.Operator.JoyBtnRaw, Cfg := cfg, NeutralXMem := nx, NeutralYMem := ny);
home(DeadmanArmed := joy.DeadmanArmed, JoystickDeflected := NOT joy.AtNeutralXY, JoystickPull := joy.AxisCmdY.DirectionPositive, JoystickPush := joy.AxisCmdY.DirectionNegative, BtnValidation := bench.Operator.JoyBtnRaw);
ASSERT_EQ(home.MachineHomingSeqStep, E_MachineHomingTxState.HX0_REPOS, 'N1/cycle : aucun HX1 par geste joystick'); ASSERT_FALSE(home.M3Locked, 'N1/cycle : aucun verrou homing parasite'); ASSERT_TRUE(home.MachineHomed, 'Reference conservee');
ADVANCE_TIME(10000000); bench(RawPosM1 := raw1, RawPosM2 := raw2);
joy(RawX := bench.Operator.JoyXRaw_ANA1, RawY := bench.Operator.JoyYRaw_ANA2, RawButton := bench.Operator.JoyBtnRaw, Cfg := cfg, NeutralXMem := nx, NeutralYMem := ny);
home(DeadmanArmed := joy.DeadmanArmed, JoystickDeflected := NOT joy.AtNeutralXY, JoystickPull := joy.AxisCmdY.DirectionPositive, JoystickPush := joy.AxisCmdY.DirectionNegative, BtnValidation := bench.Operator.JoyBtnRaw);
ASSERT_EQ(home.MachineHomingSeqStep, E_MachineHomingTxState.HX0_REPOS, 'N1/cycle : aucun HX1 par geste joystick'); ASSERT_FALSE(home.M3Locked, 'N1/cycle : aucun verrou homing parasite'); ASSERT_TRUE(home.MachineHomed, 'Reference conservee');
ADVANCE_TIME(10000000); bench(RawPosM1 := raw1, RawPosM2 := raw2);
joy(RawX := bench.Operator.JoyXRaw_ANA1, RawY := bench.Operator.JoyYRaw_ANA2, RawButton := bench.Operator.JoyBtnRaw, Cfg := cfg, NeutralXMem := nx, NeutralYMem := ny);
home(DeadmanArmed := joy.DeadmanArmed, JoystickDeflected := NOT joy.AtNeutralXY, JoystickPull := joy.AxisCmdY.DirectionPositive, JoystickPush := joy.AxisCmdY.DirectionNegative, BtnValidation := bench.Operator.JoyBtnRaw);
ASSERT_EQ(home.MachineHomingSeqStep, E_MachineHomingTxState.HX0_REPOS, 'N1/cycle : aucun HX1 par geste joystick'); ASSERT_FALSE(home.M3Locked, 'N1/cycle : aucun verrou homing parasite'); ASSERT_TRUE(home.MachineHomed, 'Reference conservee');
ADVANCE_TIME(10000000); bench(RawPosM1 := raw1, RawPosM2 := raw2);
joy(RawX := bench.Operator.JoyXRaw_ANA1, RawY := bench.Operator.JoyYRaw_ANA2, RawButton := bench.Operator.JoyBtnRaw, Cfg := cfg, NeutralXMem := nx, NeutralYMem := ny);
home(DeadmanArmed := joy.DeadmanArmed, JoystickDeflected := NOT joy.AtNeutralXY, JoystickPull := joy.AxisCmdY.DirectionPositive, JoystickPush := joy.AxisCmdY.DirectionNegative, BtnValidation := bench.Operator.JoyBtnRaw);
ASSERT_EQ(home.MachineHomingSeqStep, E_MachineHomingTxState.HX0_REPOS, 'N1/cycle : aucun HX1 par geste joystick'); ASSERT_FALSE(home.M3Locked, 'N1/cycle : aucun verrou homing parasite'); ASSERT_TRUE(home.MachineHomed, 'Reference conservee');
ADVANCE_TIME(10000000); bench(RawPosM1 := raw1, RawPosM2 := raw2);
joy(RawX := bench.Operator.JoyXRaw_ANA1, RawY := bench.Operator.JoyYRaw_ANA2, RawButton := bench.Operator.JoyBtnRaw, Cfg := cfg, NeutralXMem := nx, NeutralYMem := ny);
home(DeadmanArmed := joy.DeadmanArmed, JoystickDeflected := NOT joy.AtNeutralXY, JoystickPull := joy.AxisCmdY.DirectionPositive, JoystickPush := joy.AxisCmdY.DirectionNegative, BtnValidation := bench.Operator.JoyBtnRaw);
ASSERT_EQ(home.MachineHomingSeqStep, E_MachineHomingTxState.HX0_REPOS, 'N1/cycle : aucun HX1 par geste joystick'); ASSERT_FALSE(home.M3Locked, 'N1/cycle : aucun verrou homing parasite'); ASSERT_TRUE(home.MachineHomed, 'Reference conservee');
ADVANCE_TIME(10000000); bench(RawPosM1 := raw1, RawPosM2 := raw2);
joy(RawX := bench.Operator.JoyXRaw_ANA1, RawY := bench.Operator.JoyYRaw_ANA2, RawButton := bench.Operator.JoyBtnRaw, Cfg := cfg, NeutralXMem := nx, NeutralYMem := ny);
home(DeadmanArmed := joy.DeadmanArmed, JoystickDeflected := NOT joy.AtNeutralXY, JoystickPull := joy.AxisCmdY.DirectionPositive, JoystickPush := joy.AxisCmdY.DirectionNegative, BtnValidation := bench.Operator.JoyBtnRaw);
ASSERT_EQ(home.MachineHomingSeqStep, E_MachineHomingTxState.HX0_REPOS, 'N1/cycle : aucun HX1 par geste joystick'); ASSERT_FALSE(home.M3Locked, 'N1/cycle : aucun verrou homing parasite'); ASSERT_TRUE(home.MachineHomed, 'Reference conservee');
ADVANCE_TIME(10000000); bench(RawPosM1 := raw1, RawPosM2 := raw2);
joy(RawX := bench.Operator.JoyXRaw_ANA1, RawY := bench.Operator.JoyYRaw_ANA2, RawButton := bench.Operator.JoyBtnRaw, Cfg := cfg, NeutralXMem := nx, NeutralYMem := ny);
home(DeadmanArmed := joy.DeadmanArmed, JoystickDeflected := NOT joy.AtNeutralXY, JoystickPull := joy.AxisCmdY.DirectionPositive, JoystickPush := joy.AxisCmdY.DirectionNegative, BtnValidation := bench.Operator.JoyBtnRaw);
ASSERT_EQ(home.MachineHomingSeqStep, E_MachineHomingTxState.HX0_REPOS, 'N1/cycle : aucun HX1 par geste joystick'); ASSERT_FALSE(home.M3Locked, 'N1/cycle : aucun verrou homing parasite'); ASSERT_TRUE(home.MachineHomed, 'Reference conservee');
ADVANCE_TIME(10000000); bench(RawPosM1 := raw1, RawPosM2 := raw2);
joy(RawX := bench.Operator.JoyXRaw_ANA1, RawY := bench.Operator.JoyYRaw_ANA2, RawButton := bench.Operator.JoyBtnRaw, Cfg := cfg, NeutralXMem := nx, NeutralYMem := ny);
home(DeadmanArmed := joy.DeadmanArmed, JoystickDeflected := NOT joy.AtNeutralXY, JoystickPull := joy.AxisCmdY.DirectionPositive, JoystickPush := joy.AxisCmdY.DirectionNegative, BtnValidation := bench.Operator.JoyBtnRaw);
ASSERT_EQ(home.MachineHomingSeqStep, E_MachineHomingTxState.HX0_REPOS, 'N1/cycle : aucun HX1 par geste joystick'); ASSERT_FALSE(home.M3Locked, 'N1/cycle : aucun verrou homing parasite'); ASSERT_TRUE(home.MachineHomed, 'Reference conservee');
ADVANCE_TIME(10000000); bench(RawPosM1 := raw1, RawPosM2 := raw2);
joy(RawX := bench.Operator.JoyXRaw_ANA1, RawY := bench.Operator.JoyYRaw_ANA2, RawButton := bench.Operator.JoyBtnRaw, Cfg := cfg, NeutralXMem := nx, NeutralYMem := ny);
home(DeadmanArmed := joy.DeadmanArmed, JoystickDeflected := NOT joy.AtNeutralXY, JoystickPull := joy.AxisCmdY.DirectionPositive, JoystickPush := joy.AxisCmdY.DirectionNegative, BtnValidation := bench.Operator.JoyBtnRaw);
ASSERT_EQ(home.MachineHomingSeqStep, E_MachineHomingTxState.HX0_REPOS, 'N1/cycle : aucun HX1 par geste joystick'); ASSERT_FALSE(home.M3Locked, 'N1/cycle : aucun verrou homing parasite'); ASSERT_TRUE(home.MachineHomed, 'Reference conservee');
ADVANCE_TIME(10000000); bench(RawPosM1 := raw1, RawPosM2 := raw2);
joy(RawX := bench.Operator.JoyXRaw_ANA1, RawY := bench.Operator.JoyYRaw_ANA2, RawButton := bench.Operator.JoyBtnRaw, Cfg := cfg, NeutralXMem := nx, NeutralYMem := ny);
home(DeadmanArmed := joy.DeadmanArmed, JoystickDeflected := NOT joy.AtNeutralXY, JoystickPull := joy.AxisCmdY.DirectionPositive, JoystickPush := joy.AxisCmdY.DirectionNegative, BtnValidation := bench.Operator.JoyBtnRaw);
ASSERT_EQ(home.MachineHomingSeqStep, E_MachineHomingTxState.HX0_REPOS, 'N1/cycle : aucun HX1 par geste joystick'); ASSERT_FALSE(home.M3Locked, 'N1/cycle : aucun verrou homing parasite'); ASSERT_TRUE(home.MachineHomed, 'Reference conservee');
ADVANCE_TIME(10000000); bench(RawPosM1 := raw1, RawPosM2 := raw2);
joy(RawX := bench.Operator.JoyXRaw_ANA1, RawY := bench.Operator.JoyYRaw_ANA2, RawButton := bench.Operator.JoyBtnRaw, Cfg := cfg, NeutralXMem := nx, NeutralYMem := ny);
home(DeadmanArmed := joy.DeadmanArmed, JoystickDeflected := NOT joy.AtNeutralXY, JoystickPull := joy.AxisCmdY.DirectionPositive, JoystickPush := joy.AxisCmdY.DirectionNegative, BtnValidation := bench.Operator.JoyBtnRaw);
ASSERT_EQ(home.MachineHomingSeqStep, E_MachineHomingTxState.HX0_REPOS, 'N1/cycle : aucun HX1 par geste joystick'); ASSERT_FALSE(home.M3Locked, 'N1/cycle : aucun verrou homing parasite'); ASSERT_TRUE(home.MachineHomed, 'Reference conservee');
ADVANCE_TIME(10000000); bench(RawPosM1 := raw1, RawPosM2 := raw2);
joy(RawX := bench.Operator.JoyXRaw_ANA1, RawY := bench.Operator.JoyYRaw_ANA2, RawButton := bench.Operator.JoyBtnRaw, Cfg := cfg, NeutralXMem := nx, NeutralYMem := ny);
home(DeadmanArmed := joy.DeadmanArmed, JoystickDeflected := NOT joy.AtNeutralXY, JoystickPull := joy.AxisCmdY.DirectionPositive, JoystickPush := joy.AxisCmdY.DirectionNegative, BtnValidation := bench.Operator.JoyBtnRaw);
ASSERT_EQ(home.MachineHomingSeqStep, E_MachineHomingTxState.HX0_REPOS, 'N1/cycle : aucun HX1 par geste joystick'); ASSERT_FALSE(home.M3Locked, 'N1/cycle : aucun verrou homing parasite'); ASSERT_TRUE(home.MachineHomed, 'Reference conservee');
ADVANCE_TIME(10000000); bench(RawPosM1 := raw1, RawPosM2 := raw2);
joy(RawX := bench.Operator.JoyXRaw_ANA1, RawY := bench.Operator.JoyYRaw_ANA2, RawButton := bench.Operator.JoyBtnRaw, Cfg := cfg, NeutralXMem := nx, NeutralYMem := ny);
home(DeadmanArmed := joy.DeadmanArmed, JoystickDeflected := NOT joy.AtNeutralXY, JoystickPull := joy.AxisCmdY.DirectionPositive, JoystickPush := joy.AxisCmdY.DirectionNegative, BtnValidation := bench.Operator.JoyBtnRaw);
ASSERT_EQ(home.MachineHomingSeqStep, E_MachineHomingTxState.HX0_REPOS, 'N1/cycle : aucun HX1 par geste joystick'); ASSERT_FALSE(home.M3Locked, 'N1/cycle : aucun verrou homing parasite'); ASSERT_TRUE(home.MachineHomed, 'Reference conservee');
ADVANCE_TIME(10000000); bench(RawPosM1 := raw1, RawPosM2 := raw2);
joy(RawX := bench.Operator.JoyXRaw_ANA1, RawY := bench.Operator.JoyYRaw_ANA2, RawButton := bench.Operator.JoyBtnRaw, Cfg := cfg, NeutralXMem := nx, NeutralYMem := ny);
home(DeadmanArmed := joy.DeadmanArmed, JoystickDeflected := NOT joy.AtNeutralXY, JoystickPull := joy.AxisCmdY.DirectionPositive, JoystickPush := joy.AxisCmdY.DirectionNegative, BtnValidation := bench.Operator.JoyBtnRaw);
ASSERT_EQ(home.MachineHomingSeqStep, E_MachineHomingTxState.HX0_REPOS, 'N1/cycle : aucun HX1 par geste joystick'); ASSERT_FALSE(home.M3Locked, 'N1/cycle : aucun verrou homing parasite'); ASSERT_TRUE(home.MachineHomed, 'Reference conservee');
ADVANCE_TIME(10000000); bench(RawPosM1 := raw1, RawPosM2 := raw2);
joy(RawX := bench.Operator.JoyXRaw_ANA1, RawY := bench.Operator.JoyYRaw_ANA2, RawButton := bench.Operator.JoyBtnRaw, Cfg := cfg, NeutralXMem := nx, NeutralYMem := ny);
home(DeadmanArmed := joy.DeadmanArmed, JoystickDeflected := NOT joy.AtNeutralXY, JoystickPull := joy.AxisCmdY.DirectionPositive, JoystickPush := joy.AxisCmdY.DirectionNegative, BtnValidation := bench.Operator.JoyBtnRaw);
ASSERT_EQ(home.MachineHomingSeqStep, E_MachineHomingTxState.HX0_REPOS, 'N1/cycle : aucun HX1 par geste joystick'); ASSERT_FALSE(home.M3Locked, 'N1/cycle : aucun verrou homing parasite'); ASSERT_TRUE(home.MachineHomed, 'Reference conservee');
ADVANCE_TIME(10000000); bench(RawPosM1 := raw1, RawPosM2 := raw2);
joy(RawX := bench.Operator.JoyXRaw_ANA1, RawY := bench.Operator.JoyYRaw_ANA2, RawButton := bench.Operator.JoyBtnRaw, Cfg := cfg, NeutralXMem := nx, NeutralYMem := ny);
home(DeadmanArmed := joy.DeadmanArmed, JoystickDeflected := NOT joy.AtNeutralXY, JoystickPull := joy.AxisCmdY.DirectionPositive, JoystickPush := joy.AxisCmdY.DirectionNegative, BtnValidation := bench.Operator.JoyBtnRaw);
ASSERT_EQ(home.MachineHomingSeqStep, E_MachineHomingTxState.HX0_REPOS, 'N1/cycle : aucun HX1 par geste joystick'); ASSERT_FALSE(home.M3Locked, 'N1/cycle : aucun verrou homing parasite'); ASSERT_TRUE(home.MachineHomed, 'Reference conservee');
ADVANCE_TIME(10000000); bench(RawPosM1 := raw1, RawPosM2 := raw2);
joy(RawX := bench.Operator.JoyXRaw_ANA1, RawY := bench.Operator.JoyYRaw_ANA2, RawButton := bench.Operator.JoyBtnRaw, Cfg := cfg, NeutralXMem := nx, NeutralYMem := ny);
home(DeadmanArmed := joy.DeadmanArmed, JoystickDeflected := NOT joy.AtNeutralXY, JoystickPull := joy.AxisCmdY.DirectionPositive, JoystickPush := joy.AxisCmdY.DirectionNegative, BtnValidation := bench.Operator.JoyBtnRaw);
ASSERT_EQ(home.MachineHomingSeqStep, E_MachineHomingTxState.HX0_REPOS, 'N1/cycle : aucun HX1 par geste joystick'); ASSERT_FALSE(home.M3Locked, 'N1/cycle : aucun verrou homing parasite'); ASSERT_TRUE(home.MachineHomed, 'Reference conservee');
ADVANCE_TIME(10000000); bench(RawPosM1 := raw1, RawPosM2 := raw2);
joy(RawX := bench.Operator.JoyXRaw_ANA1, RawY := bench.Operator.JoyYRaw_ANA2, RawButton := bench.Operator.JoyBtnRaw, Cfg := cfg, NeutralXMem := nx, NeutralYMem := ny);
home(DeadmanArmed := joy.DeadmanArmed, JoystickDeflected := NOT joy.AtNeutralXY, JoystickPull := joy.AxisCmdY.DirectionPositive, JoystickPush := joy.AxisCmdY.DirectionNegative, BtnValidation := bench.Operator.JoyBtnRaw);
ASSERT_EQ(home.MachineHomingSeqStep, E_MachineHomingTxState.HX0_REPOS, 'N1/cycle : aucun HX1 par geste joystick'); ASSERT_FALSE(home.M3Locked, 'N1/cycle : aucun verrou homing parasite'); ASSERT_TRUE(home.MachineHomed, 'Reference conservee');
ADVANCE_TIME(10000000); bench(RawPosM1 := raw1, RawPosM2 := raw2);
joy(RawX := bench.Operator.JoyXRaw_ANA1, RawY := bench.Operator.JoyYRaw_ANA2, RawButton := bench.Operator.JoyBtnRaw, Cfg := cfg, NeutralXMem := nx, NeutralYMem := ny);
home(DeadmanArmed := joy.DeadmanArmed, JoystickDeflected := NOT joy.AtNeutralXY, JoystickPull := joy.AxisCmdY.DirectionPositive, JoystickPush := joy.AxisCmdY.DirectionNegative, BtnValidation := bench.Operator.JoyBtnRaw);
ASSERT_EQ(home.MachineHomingSeqStep, E_MachineHomingTxState.HX0_REPOS, 'N1/cycle : aucun HX1 par geste joystick'); ASSERT_FALSE(home.M3Locked, 'N1/cycle : aucun verrou homing parasite'); ASSERT_TRUE(home.MachineHomed, 'Reference conservee');
ADVANCE_TIME(10000000); bench(RawPosM1 := raw1, RawPosM2 := raw2);
joy(RawX := bench.Operator.JoyXRaw_ANA1, RawY := bench.Operator.JoyYRaw_ANA2, RawButton := bench.Operator.JoyBtnRaw, Cfg := cfg, NeutralXMem := nx, NeutralYMem := ny);
home(DeadmanArmed := joy.DeadmanArmed, JoystickDeflected := NOT joy.AtNeutralXY, JoystickPull := joy.AxisCmdY.DirectionPositive, JoystickPush := joy.AxisCmdY.DirectionNegative, BtnValidation := bench.Operator.JoyBtnRaw);
ASSERT_EQ(home.MachineHomingSeqStep, E_MachineHomingTxState.HX0_REPOS, 'N1/cycle : aucun HX1 par geste joystick'); ASSERT_FALSE(home.M3Locked, 'N1/cycle : aucun verrou homing parasite'); ASSERT_TRUE(home.MachineHomed, 'Reference conservee');
ADVANCE_TIME(10000000); bench(RawPosM1 := raw1, RawPosM2 := raw2);
joy(RawX := bench.Operator.JoyXRaw_ANA1, RawY := bench.Operator.JoyYRaw_ANA2, RawButton := bench.Operator.JoyBtnRaw, Cfg := cfg, NeutralXMem := nx, NeutralYMem := ny);
home(DeadmanArmed := joy.DeadmanArmed, JoystickDeflected := NOT joy.AtNeutralXY, JoystickPull := joy.AxisCmdY.DirectionPositive, JoystickPush := joy.AxisCmdY.DirectionNegative, BtnValidation := bench.Operator.JoyBtnRaw);
ASSERT_EQ(home.MachineHomingSeqStep, E_MachineHomingTxState.HX0_REPOS, 'N1/cycle : aucun HX1 par geste joystick'); ASSERT_FALSE(home.M3Locked, 'N1/cycle : aucun verrou homing parasite'); ASSERT_TRUE(home.MachineHomed, 'Reference conservee');
ADVANCE_TIME(10000000); bench(RawPosM1 := raw1, RawPosM2 := raw2);
joy(RawX := bench.Operator.JoyXRaw_ANA1, RawY := bench.Operator.JoyYRaw_ANA2, RawButton := bench.Operator.JoyBtnRaw, Cfg := cfg, NeutralXMem := nx, NeutralYMem := ny);
home(DeadmanArmed := joy.DeadmanArmed, JoystickDeflected := NOT joy.AtNeutralXY, JoystickPull := joy.AxisCmdY.DirectionPositive, JoystickPush := joy.AxisCmdY.DirectionNegative, BtnValidation := bench.Operator.JoyBtnRaw);
ASSERT_EQ(home.MachineHomingSeqStep, E_MachineHomingTxState.HX0_REPOS, 'N1/cycle : aucun HX1 par geste joystick'); ASSERT_FALSE(home.M3Locked, 'N1/cycle : aucun verrou homing parasite'); ASSERT_TRUE(home.MachineHomed, 'Reference conservee');
ADVANCE_TIME(10000000); bench(RawPosM1 := raw1, RawPosM2 := raw2);
joy(RawX := bench.Operator.JoyXRaw_ANA1, RawY := bench.Operator.JoyYRaw_ANA2, RawButton := bench.Operator.JoyBtnRaw, Cfg := cfg, NeutralXMem := nx, NeutralYMem := ny);
home(DeadmanArmed := joy.DeadmanArmed, JoystickDeflected := NOT joy.AtNeutralXY, JoystickPull := joy.AxisCmdY.DirectionPositive, JoystickPush := joy.AxisCmdY.DirectionNegative, BtnValidation := bench.Operator.JoyBtnRaw);
ASSERT_EQ(home.MachineHomingSeqStep, E_MachineHomingTxState.HX0_REPOS, 'N1/cycle : aucun HX1 par geste joystick'); ASSERT_FALSE(home.M3Locked, 'N1/cycle : aucun verrou homing parasite'); ASSERT_TRUE(home.MachineHomed, 'Reference conservee');
ADVANCE_TIME(10000000); bench(RawPosM1 := raw1, RawPosM2 := raw2);
joy(RawX := bench.Operator.JoyXRaw_ANA1, RawY := bench.Operator.JoyYRaw_ANA2, RawButton := bench.Operator.JoyBtnRaw, Cfg := cfg, NeutralXMem := nx, NeutralYMem := ny);
home(DeadmanArmed := joy.DeadmanArmed, JoystickDeflected := NOT joy.AtNeutralXY, JoystickPull := joy.AxisCmdY.DirectionPositive, JoystickPush := joy.AxisCmdY.DirectionNegative, BtnValidation := bench.Operator.JoyBtnRaw);
ASSERT_EQ(home.MachineHomingSeqStep, E_MachineHomingTxState.HX0_REPOS, 'N1/cycle : aucun HX1 par geste joystick'); ASSERT_FALSE(home.M3Locked, 'N1/cycle : aucun verrou homing parasite'); ASSERT_TRUE(home.MachineHomed, 'Reference conservee');
ADVANCE_TIME(10000000); bench(RawPosM1 := raw1, RawPosM2 := raw2);
joy(RawX := bench.Operator.JoyXRaw_ANA1, RawY := bench.Operator.JoyYRaw_ANA2, RawButton := bench.Operator.JoyBtnRaw, Cfg := cfg, NeutralXMem := nx, NeutralYMem := ny);
home(DeadmanArmed := joy.DeadmanArmed, JoystickDeflected := NOT joy.AtNeutralXY, JoystickPull := joy.AxisCmdY.DirectionPositive, JoystickPush := joy.AxisCmdY.DirectionNegative, BtnValidation := bench.Operator.JoyBtnRaw);
ASSERT_EQ(home.MachineHomingSeqStep, E_MachineHomingTxState.HX0_REPOS, 'N1/cycle : aucun HX1 par geste joystick'); ASSERT_FALSE(home.M3Locked, 'N1/cycle : aucun verrou homing parasite'); ASSERT_TRUE(home.MachineHomed, 'Reference conservee');
ADVANCE_TIME(10000000); bench(RawPosM1 := raw1, RawPosM2 := raw2);
joy(RawX := bench.Operator.JoyXRaw_ANA1, RawY := bench.Operator.JoyYRaw_ANA2, RawButton := bench.Operator.JoyBtnRaw, Cfg := cfg, NeutralXMem := nx, NeutralYMem := ny);
home(DeadmanArmed := joy.DeadmanArmed, JoystickDeflected := NOT joy.AtNeutralXY, JoystickPull := joy.AxisCmdY.DirectionPositive, JoystickPush := joy.AxisCmdY.DirectionNegative, BtnValidation := bench.Operator.JoyBtnRaw);
ASSERT_EQ(home.MachineHomingSeqStep, E_MachineHomingTxState.HX0_REPOS, 'N1/cycle : aucun HX1 par geste joystick'); ASSERT_FALSE(home.M3Locked, 'N1/cycle : aucun verrou homing parasite'); ASSERT_TRUE(home.MachineHomed, 'Reference conservee');
ADVANCE_TIME(10000000); bench(RawPosM1 := raw1, RawPosM2 := raw2);
joy(RawX := bench.Operator.JoyXRaw_ANA1, RawY := bench.Operator.JoyYRaw_ANA2, RawButton := bench.Operator.JoyBtnRaw, Cfg := cfg, NeutralXMem := nx, NeutralYMem := ny);
home(DeadmanArmed := joy.DeadmanArmed, JoystickDeflected := NOT joy.AtNeutralXY, JoystickPull := joy.AxisCmdY.DirectionPositive, JoystickPush := joy.AxisCmdY.DirectionNegative, BtnValidation := bench.Operator.JoyBtnRaw);
ASSERT_EQ(home.MachineHomingSeqStep, E_MachineHomingTxState.HX0_REPOS, 'N1/cycle : aucun HX1 par geste joystick'); ASSERT_FALSE(home.M3Locked, 'N1/cycle : aucun verrou homing parasite'); ASSERT_TRUE(home.MachineHomed, 'Reference conservee');
ADVANCE_TIME(10000000); bench(RawPosM1 := raw1, RawPosM2 := raw2);
joy(RawX := bench.Operator.JoyXRaw_ANA1, RawY := bench.Operator.JoyYRaw_ANA2, RawButton := bench.Operator.JoyBtnRaw, Cfg := cfg, NeutralXMem := nx, NeutralYMem := ny);
home(DeadmanArmed := joy.DeadmanArmed, JoystickDeflected := NOT joy.AtNeutralXY, JoystickPull := joy.AxisCmdY.DirectionPositive, JoystickPush := joy.AxisCmdY.DirectionNegative, BtnValidation := bench.Operator.JoyBtnRaw);
ASSERT_EQ(home.MachineHomingSeqStep, E_MachineHomingTxState.HX0_REPOS, 'N1/cycle : aucun HX1 par geste joystick'); ASSERT_FALSE(home.M3Locked, 'N1/cycle : aucun verrou homing parasite'); ASSERT_TRUE(home.MachineHomed, 'Reference conservee');
ADVANCE_TIME(10000000); bench(RawPosM1 := raw1, RawPosM2 := raw2);
joy(RawX := bench.Operator.JoyXRaw_ANA1, RawY := bench.Operator.JoyYRaw_ANA2, RawButton := bench.Operator.JoyBtnRaw, Cfg := cfg, NeutralXMem := nx, NeutralYMem := ny);
home(DeadmanArmed := joy.DeadmanArmed, JoystickDeflected := NOT joy.AtNeutralXY, JoystickPull := joy.AxisCmdY.DirectionPositive, JoystickPush := joy.AxisCmdY.DirectionNegative, BtnValidation := bench.Operator.JoyBtnRaw);
ASSERT_EQ(home.MachineHomingSeqStep, E_MachineHomingTxState.HX0_REPOS, 'N1/cycle : aucun HX1 par geste joystick'); ASSERT_FALSE(home.M3Locked, 'N1/cycle : aucun verrou homing parasite'); ASSERT_TRUE(home.MachineHomed, 'Reference conservee');
ASSERT_TRUE(joy.AxisCmdY.DirectionNegative, 'Geste joystick en mode cycle disponible');
bench.SimJoystickRev_Down_Open_Active := FALSE;
ADVANCE_TIME(10000000); bench(RawPosM1 := raw1, RawPosM2 := raw2);
joy(RawX := bench.Operator.JoyXRaw_ANA1, RawY := bench.Operator.JoyYRaw_ANA2, RawButton := bench.Operator.JoyBtnRaw, Cfg := cfg, NeutralXMem := nx, NeutralYMem := ny);
home(DeadmanArmed := joy.DeadmanArmed, JoystickDeflected := NOT joy.AtNeutralXY, JoystickPull := joy.AxisCmdY.DirectionPositive, JoystickPush := joy.AxisCmdY.DirectionNegative, BtnValidation := bench.Operator.JoyBtnRaw);
ASSERT_EQ(home.MachineHomingSeqStep, E_MachineHomingTxState.HX0_REPOS, 'N1/cycle : aucun HX1 par geste joystick'); ASSERT_FALSE(home.M3Locked, 'N1/cycle : aucun verrou homing parasite'); ASSERT_TRUE(home.MachineHomed, 'Reference conservee');
ADVANCE_TIME(10000000); bench(RawPosM1 := raw1, RawPosM2 := raw2);
joy(RawX := bench.Operator.JoyXRaw_ANA1, RawY := bench.Operator.JoyYRaw_ANA2, RawButton := bench.Operator.JoyBtnRaw, Cfg := cfg, NeutralXMem := nx, NeutralYMem := ny);
home(DeadmanArmed := joy.DeadmanArmed, JoystickDeflected := NOT joy.AtNeutralXY, JoystickPull := joy.AxisCmdY.DirectionPositive, JoystickPush := joy.AxisCmdY.DirectionNegative, BtnValidation := bench.Operator.JoyBtnRaw);
ASSERT_EQ(home.MachineHomingSeqStep, E_MachineHomingTxState.HX0_REPOS, 'N1/cycle : aucun HX1 par geste joystick'); ASSERT_FALSE(home.M3Locked, 'N1/cycle : aucun verrou homing parasite'); ASSERT_TRUE(home.MachineHomed, 'Reference conservee');
ADVANCE_TIME(10000000); bench(RawPosM1 := raw1, RawPosM2 := raw2);
joy(RawX := bench.Operator.JoyXRaw_ANA1, RawY := bench.Operator.JoyYRaw_ANA2, RawButton := bench.Operator.JoyBtnRaw, Cfg := cfg, NeutralXMem := nx, NeutralYMem := ny);
home(DeadmanArmed := joy.DeadmanArmed, JoystickDeflected := NOT joy.AtNeutralXY, JoystickPull := joy.AxisCmdY.DirectionPositive, JoystickPush := joy.AxisCmdY.DirectionNegative, BtnValidation := bench.Operator.JoyBtnRaw);
ASSERT_EQ(home.MachineHomingSeqStep, E_MachineHomingTxState.HX0_REPOS, 'N1/cycle : aucun HX1 par geste joystick'); ASSERT_FALSE(home.M3Locked, 'N1/cycle : aucun verrou homing parasite'); ASSERT_TRUE(home.MachineHomed, 'Reference conservee');
ADVANCE_TIME(10000000); bench(RawPosM1 := raw1, RawPosM2 := raw2);
joy(RawX := bench.Operator.JoyXRaw_ANA1, RawY := bench.Operator.JoyYRaw_ANA2, RawButton := bench.Operator.JoyBtnRaw, Cfg := cfg, NeutralXMem := nx, NeutralYMem := ny);
home(DeadmanArmed := joy.DeadmanArmed, JoystickDeflected := NOT joy.AtNeutralXY, JoystickPull := joy.AxisCmdY.DirectionPositive, JoystickPush := joy.AxisCmdY.DirectionNegative, BtnValidation := bench.Operator.JoyBtnRaw);
ASSERT_EQ(home.MachineHomingSeqStep, E_MachineHomingTxState.HX0_REPOS, 'N1/cycle : aucun HX1 par geste joystick'); ASSERT_FALSE(home.M3Locked, 'N1/cycle : aucun verrou homing parasite'); ASSERT_TRUE(home.MachineHomed, 'Reference conservee');
ADVANCE_TIME(10000000); bench(RawPosM1 := raw1, RawPosM2 := raw2);
joy(RawX := bench.Operator.JoyXRaw_ANA1, RawY := bench.Operator.JoyYRaw_ANA2, RawButton := bench.Operator.JoyBtnRaw, Cfg := cfg, NeutralXMem := nx, NeutralYMem := ny);
home(DeadmanArmed := joy.DeadmanArmed, JoystickDeflected := NOT joy.AtNeutralXY, JoystickPull := joy.AxisCmdY.DirectionPositive, JoystickPush := joy.AxisCmdY.DirectionNegative, BtnValidation := bench.Operator.JoyBtnRaw);
ASSERT_EQ(home.MachineHomingSeqStep, E_MachineHomingTxState.HX0_REPOS, 'N1/cycle : aucun HX1 par geste joystick'); ASSERT_FALSE(home.M3Locked, 'N1/cycle : aucun verrou homing parasite'); ASSERT_TRUE(home.MachineHomed, 'Reference conservee');
ADVANCE_TIME(10000000); bench(RawPosM1 := raw1, RawPosM2 := raw2);
joy(RawX := bench.Operator.JoyXRaw_ANA1, RawY := bench.Operator.JoyYRaw_ANA2, RawButton := bench.Operator.JoyBtnRaw, Cfg := cfg, NeutralXMem := nx, NeutralYMem := ny);
home(DeadmanArmed := joy.DeadmanArmed, JoystickDeflected := NOT joy.AtNeutralXY, JoystickPull := joy.AxisCmdY.DirectionPositive, JoystickPush := joy.AxisCmdY.DirectionNegative, BtnValidation := bench.Operator.JoyBtnRaw);
ASSERT_EQ(home.MachineHomingSeqStep, E_MachineHomingTxState.HX0_REPOS, 'N1/cycle : aucun HX1 par geste joystick'); ASSERT_FALSE(home.M3Locked, 'N1/cycle : aucun verrou homing parasite'); ASSERT_TRUE(home.MachineHomed, 'Reference conservee');
ADVANCE_TIME(10000000); bench(RawPosM1 := raw1, RawPosM2 := raw2);
joy(RawX := bench.Operator.JoyXRaw_ANA1, RawY := bench.Operator.JoyYRaw_ANA2, RawButton := bench.Operator.JoyBtnRaw, Cfg := cfg, NeutralXMem := nx, NeutralYMem := ny);
home(DeadmanArmed := joy.DeadmanArmed, JoystickDeflected := NOT joy.AtNeutralXY, JoystickPull := joy.AxisCmdY.DirectionPositive, JoystickPush := joy.AxisCmdY.DirectionNegative, BtnValidation := bench.Operator.JoyBtnRaw);
ASSERT_EQ(home.MachineHomingSeqStep, E_MachineHomingTxState.HX0_REPOS, 'N1/cycle : aucun HX1 par geste joystick'); ASSERT_FALSE(home.M3Locked, 'N1/cycle : aucun verrou homing parasite'); ASSERT_TRUE(home.MachineHomed, 'Reference conservee');
ADVANCE_TIME(10000000); bench(RawPosM1 := raw1, RawPosM2 := raw2);
joy(RawX := bench.Operator.JoyXRaw_ANA1, RawY := bench.Operator.JoyYRaw_ANA2, RawButton := bench.Operator.JoyBtnRaw, Cfg := cfg, NeutralXMem := nx, NeutralYMem := ny);
home(DeadmanArmed := joy.DeadmanArmed, JoystickDeflected := NOT joy.AtNeutralXY, JoystickPull := joy.AxisCmdY.DirectionPositive, JoystickPush := joy.AxisCmdY.DirectionNegative, BtnValidation := bench.Operator.JoyBtnRaw);
ASSERT_EQ(home.MachineHomingSeqStep, E_MachineHomingTxState.HX0_REPOS, 'N1/cycle : aucun HX1 par geste joystick'); ASSERT_FALSE(home.M3Locked, 'N1/cycle : aucun verrou homing parasite'); ASSERT_TRUE(home.MachineHomed, 'Reference conservee');
ADVANCE_TIME(10000000); bench(RawPosM1 := raw1, RawPosM2 := raw2);
joy(RawX := bench.Operator.JoyXRaw_ANA1, RawY := bench.Operator.JoyYRaw_ANA2, RawButton := bench.Operator.JoyBtnRaw, Cfg := cfg, NeutralXMem := nx, NeutralYMem := ny);
home(DeadmanArmed := joy.DeadmanArmed, JoystickDeflected := NOT joy.AtNeutralXY, JoystickPull := joy.AxisCmdY.DirectionPositive, JoystickPush := joy.AxisCmdY.DirectionNegative, BtnValidation := bench.Operator.JoyBtnRaw);
ASSERT_EQ(home.MachineHomingSeqStep, E_MachineHomingTxState.HX0_REPOS, 'N1/cycle : aucun HX1 par geste joystick'); ASSERT_FALSE(home.M3Locked, 'N1/cycle : aucun verrou homing parasite'); ASSERT_TRUE(home.MachineHomed, 'Reference conservee');
ADVANCE_TIME(10000000); bench(RawPosM1 := raw1, RawPosM2 := raw2);
joy(RawX := bench.Operator.JoyXRaw_ANA1, RawY := bench.Operator.JoyYRaw_ANA2, RawButton := bench.Operator.JoyBtnRaw, Cfg := cfg, NeutralXMem := nx, NeutralYMem := ny);
home(DeadmanArmed := joy.DeadmanArmed, JoystickDeflected := NOT joy.AtNeutralXY, JoystickPull := joy.AxisCmdY.DirectionPositive, JoystickPush := joy.AxisCmdY.DirectionNegative, BtnValidation := bench.Operator.JoyBtnRaw);
ASSERT_EQ(home.MachineHomingSeqStep, E_MachineHomingTxState.HX0_REPOS, 'N1/cycle : aucun HX1 par geste joystick'); ASSERT_FALSE(home.M3Locked, 'N1/cycle : aucun verrou homing parasite'); ASSERT_TRUE(home.MachineHomed, 'Reference conservee');
ADVANCE_TIME(10000000); bench(RawPosM1 := raw1, RawPosM2 := raw2);
joy(RawX := bench.Operator.JoyXRaw_ANA1, RawY := bench.Operator.JoyYRaw_ANA2, RawButton := bench.Operator.JoyBtnRaw, Cfg := cfg, NeutralXMem := nx, NeutralYMem := ny);
home(DeadmanArmed := joy.DeadmanArmed, JoystickDeflected := NOT joy.AtNeutralXY, JoystickPull := joy.AxisCmdY.DirectionPositive, JoystickPush := joy.AxisCmdY.DirectionNegative, BtnValidation := bench.Operator.JoyBtnRaw);
ASSERT_EQ(home.MachineHomingSeqStep, E_MachineHomingTxState.HX0_REPOS, 'N1/cycle : aucun HX1 par geste joystick'); ASSERT_FALSE(home.M3Locked, 'N1/cycle : aucun verrou homing parasite'); ASSERT_TRUE(home.MachineHomed, 'Reference conservee');
ADVANCE_TIME(10000000); bench(RawPosM1 := raw1, RawPosM2 := raw2);
joy(RawX := bench.Operator.JoyXRaw_ANA1, RawY := bench.Operator.JoyYRaw_ANA2, RawButton := bench.Operator.JoyBtnRaw, Cfg := cfg, NeutralXMem := nx, NeutralYMem := ny);
home(DeadmanArmed := joy.DeadmanArmed, JoystickDeflected := NOT joy.AtNeutralXY, JoystickPull := joy.AxisCmdY.DirectionPositive, JoystickPush := joy.AxisCmdY.DirectionNegative, BtnValidation := bench.Operator.JoyBtnRaw);
ASSERT_EQ(home.MachineHomingSeqStep, E_MachineHomingTxState.HX0_REPOS, 'N1/cycle : aucun HX1 par geste joystick'); ASSERT_FALSE(home.M3Locked, 'N1/cycle : aucun verrou homing parasite'); ASSERT_TRUE(home.MachineHomed, 'Reference conservee');
ADVANCE_TIME(10000000); bench(RawPosM1 := raw1, RawPosM2 := raw2);
joy(RawX := bench.Operator.JoyXRaw_ANA1, RawY := bench.Operator.JoyYRaw_ANA2, RawButton := bench.Operator.JoyBtnRaw, Cfg := cfg, NeutralXMem := nx, NeutralYMem := ny);
home(DeadmanArmed := joy.DeadmanArmed, JoystickDeflected := NOT joy.AtNeutralXY, JoystickPull := joy.AxisCmdY.DirectionPositive, JoystickPush := joy.AxisCmdY.DirectionNegative, BtnValidation := bench.Operator.JoyBtnRaw);
ASSERT_EQ(home.MachineHomingSeqStep, E_MachineHomingTxState.HX0_REPOS, 'N1/cycle : aucun HX1 par geste joystick'); ASSERT_FALSE(home.M3Locked, 'N1/cycle : aucun verrou homing parasite'); ASSERT_TRUE(home.MachineHomed, 'Reference conservee');
ADVANCE_TIME(10000000); bench(RawPosM1 := raw1, RawPosM2 := raw2);
joy(RawX := bench.Operator.JoyXRaw_ANA1, RawY := bench.Operator.JoyYRaw_ANA2, RawButton := bench.Operator.JoyBtnRaw, Cfg := cfg, NeutralXMem := nx, NeutralYMem := ny);
home(DeadmanArmed := joy.DeadmanArmed, JoystickDeflected := NOT joy.AtNeutralXY, JoystickPull := joy.AxisCmdY.DirectionPositive, JoystickPush := joy.AxisCmdY.DirectionNegative, BtnValidation := bench.Operator.JoyBtnRaw);
ASSERT_EQ(home.MachineHomingSeqStep, E_MachineHomingTxState.HX0_REPOS, 'N1/cycle : aucun HX1 par geste joystick'); ASSERT_FALSE(home.M3Locked, 'N1/cycle : aucun verrou homing parasite'); ASSERT_TRUE(home.MachineHomed, 'Reference conservee');
ADVANCE_TIME(10000000); bench(RawPosM1 := raw1, RawPosM2 := raw2);
joy(RawX := bench.Operator.JoyXRaw_ANA1, RawY := bench.Operator.JoyYRaw_ANA2, RawButton := bench.Operator.JoyBtnRaw, Cfg := cfg, NeutralXMem := nx, NeutralYMem := ny);
home(DeadmanArmed := joy.DeadmanArmed, JoystickDeflected := NOT joy.AtNeutralXY, JoystickPull := joy.AxisCmdY.DirectionPositive, JoystickPush := joy.AxisCmdY.DirectionNegative, BtnValidation := bench.Operator.JoyBtnRaw);
ASSERT_EQ(home.MachineHomingSeqStep, E_MachineHomingTxState.HX0_REPOS, 'N1/cycle : aucun HX1 par geste joystick'); ASSERT_FALSE(home.M3Locked, 'N1/cycle : aucun verrou homing parasite'); ASSERT_TRUE(home.MachineHomed, 'Reference conservee');
ADVANCE_TIME(10000000); bench(RawPosM1 := raw1, RawPosM2 := raw2);
joy(RawX := bench.Operator.JoyXRaw_ANA1, RawY := bench.Operator.JoyYRaw_ANA2, RawButton := bench.Operator.JoyBtnRaw, Cfg := cfg, NeutralXMem := nx, NeutralYMem := ny);
home(DeadmanArmed := joy.DeadmanArmed, JoystickDeflected := NOT joy.AtNeutralXY, JoystickPull := joy.AxisCmdY.DirectionPositive, JoystickPush := joy.AxisCmdY.DirectionNegative, BtnValidation := bench.Operator.JoyBtnRaw);
ASSERT_EQ(home.MachineHomingSeqStep, E_MachineHomingTxState.HX0_REPOS, 'N1/cycle : aucun HX1 par geste joystick'); ASSERT_FALSE(home.M3Locked, 'N1/cycle : aucun verrou homing parasite'); ASSERT_TRUE(home.MachineHomed, 'Reference conservee');
ADVANCE_TIME(10000000); bench(RawPosM1 := raw1, RawPosM2 := raw2);
joy(RawX := bench.Operator.JoyXRaw_ANA1, RawY := bench.Operator.JoyYRaw_ANA2, RawButton := bench.Operator.JoyBtnRaw, Cfg := cfg, NeutralXMem := nx, NeutralYMem := ny);
home(DeadmanArmed := joy.DeadmanArmed, JoystickDeflected := NOT joy.AtNeutralXY, JoystickPull := joy.AxisCmdY.DirectionPositive, JoystickPush := joy.AxisCmdY.DirectionNegative, BtnValidation := bench.Operator.JoyBtnRaw);
ASSERT_EQ(home.MachineHomingSeqStep, E_MachineHomingTxState.HX0_REPOS, 'N1/cycle : aucun HX1 par geste joystick'); ASSERT_FALSE(home.M3Locked, 'N1/cycle : aucun verrou homing parasite'); ASSERT_TRUE(home.MachineHomed, 'Reference conservee');
ADVANCE_TIME(10000000); bench(RawPosM1 := raw1, RawPosM2 := raw2);
joy(RawX := bench.Operator.JoyXRaw_ANA1, RawY := bench.Operator.JoyYRaw_ANA2, RawButton := bench.Operator.JoyBtnRaw, Cfg := cfg, NeutralXMem := nx, NeutralYMem := ny);
home(DeadmanArmed := joy.DeadmanArmed, JoystickDeflected := NOT joy.AtNeutralXY, JoystickPull := joy.AxisCmdY.DirectionPositive, JoystickPush := joy.AxisCmdY.DirectionNegative, BtnValidation := bench.Operator.JoyBtnRaw);
ASSERT_EQ(home.MachineHomingSeqStep, E_MachineHomingTxState.HX0_REPOS, 'N1/cycle : aucun HX1 par geste joystick'); ASSERT_FALSE(home.M3Locked, 'N1/cycle : aucun verrou homing parasite'); ASSERT_TRUE(home.MachineHomed, 'Reference conservee');
ADVANCE_TIME(10000000); bench(RawPosM1 := raw1, RawPosM2 := raw2);
joy(RawX := bench.Operator.JoyXRaw_ANA1, RawY := bench.Operator.JoyYRaw_ANA2, RawButton := bench.Operator.JoyBtnRaw, Cfg := cfg, NeutralXMem := nx, NeutralYMem := ny);
home(DeadmanArmed := joy.DeadmanArmed, JoystickDeflected := NOT joy.AtNeutralXY, JoystickPull := joy.AxisCmdY.DirectionPositive, JoystickPush := joy.AxisCmdY.DirectionNegative, BtnValidation := bench.Operator.JoyBtnRaw);
ASSERT_EQ(home.MachineHomingSeqStep, E_MachineHomingTxState.HX0_REPOS, 'N1/cycle : aucun HX1 par geste joystick'); ASSERT_FALSE(home.M3Locked, 'N1/cycle : aucun verrou homing parasite'); ASSERT_TRUE(home.MachineHomed, 'Reference conservee');
ADVANCE_TIME(10000000); bench(RawPosM1 := raw1, RawPosM2 := raw2);
joy(RawX := bench.Operator.JoyXRaw_ANA1, RawY := bench.Operator.JoyYRaw_ANA2, RawButton := bench.Operator.JoyBtnRaw, Cfg := cfg, NeutralXMem := nx, NeutralYMem := ny);
home(DeadmanArmed := joy.DeadmanArmed, JoystickDeflected := NOT joy.AtNeutralXY, JoystickPull := joy.AxisCmdY.DirectionPositive, JoystickPush := joy.AxisCmdY.DirectionNegative, BtnValidation := bench.Operator.JoyBtnRaw);
ASSERT_EQ(home.MachineHomingSeqStep, E_MachineHomingTxState.HX0_REPOS, 'N1/cycle : aucun HX1 par geste joystick'); ASSERT_FALSE(home.M3Locked, 'N1/cycle : aucun verrou homing parasite'); ASSERT_TRUE(home.MachineHomed, 'Reference conservee');
ADVANCE_TIME(10000000); bench(RawPosM1 := raw1, RawPosM2 := raw2);
joy(RawX := bench.Operator.JoyXRaw_ANA1, RawY := bench.Operator.JoyYRaw_ANA2, RawButton := bench.Operator.JoyBtnRaw, Cfg := cfg, NeutralXMem := nx, NeutralYMem := ny);
home(DeadmanArmed := joy.DeadmanArmed, JoystickDeflected := NOT joy.AtNeutralXY, JoystickPull := joy.AxisCmdY.DirectionPositive, JoystickPush := joy.AxisCmdY.DirectionNegative, BtnValidation := bench.Operator.JoyBtnRaw);
ASSERT_EQ(home.MachineHomingSeqStep, E_MachineHomingTxState.HX0_REPOS, 'N1/cycle : aucun HX1 par geste joystick'); ASSERT_FALSE(home.M3Locked, 'N1/cycle : aucun verrou homing parasite'); ASSERT_TRUE(home.MachineHomed, 'Reference conservee');
ADVANCE_TIME(10000000); bench(RawPosM1 := raw1, RawPosM2 := raw2);
joy(RawX := bench.Operator.JoyXRaw_ANA1, RawY := bench.Operator.JoyYRaw_ANA2, RawButton := bench.Operator.JoyBtnRaw, Cfg := cfg, NeutralXMem := nx, NeutralYMem := ny);
home(DeadmanArmed := joy.DeadmanArmed, JoystickDeflected := NOT joy.AtNeutralXY, JoystickPull := joy.AxisCmdY.DirectionPositive, JoystickPush := joy.AxisCmdY.DirectionNegative, BtnValidation := bench.Operator.JoyBtnRaw);
ASSERT_EQ(home.MachineHomingSeqStep, E_MachineHomingTxState.HX0_REPOS, 'N1/cycle : aucun HX1 par geste joystick'); ASSERT_FALSE(home.M3Locked, 'N1/cycle : aucun verrou homing parasite'); ASSERT_TRUE(home.MachineHomed, 'Reference conservee');
ADVANCE_TIME(10000000); bench(RawPosM1 := raw1, RawPosM2 := raw2);
joy(RawX := bench.Operator.JoyXRaw_ANA1, RawY := bench.Operator.JoyYRaw_ANA2, RawButton := bench.Operator.JoyBtnRaw, Cfg := cfg, NeutralXMem := nx, NeutralYMem := ny);
home(DeadmanArmed := joy.DeadmanArmed, JoystickDeflected := NOT joy.AtNeutralXY, JoystickPull := joy.AxisCmdY.DirectionPositive, JoystickPush := joy.AxisCmdY.DirectionNegative, BtnValidation := bench.Operator.JoyBtnRaw);
ASSERT_EQ(home.MachineHomingSeqStep, E_MachineHomingTxState.HX0_REPOS, 'N1/cycle : aucun HX1 par geste joystick'); ASSERT_FALSE(home.M3Locked, 'N1/cycle : aucun verrou homing parasite'); ASSERT_TRUE(home.MachineHomed, 'Reference conservee');
ADVANCE_TIME(10000000); bench(RawPosM1 := raw1, RawPosM2 := raw2);
joy(RawX := bench.Operator.JoyXRaw_ANA1, RawY := bench.Operator.JoyYRaw_ANA2, RawButton := bench.Operator.JoyBtnRaw, Cfg := cfg, NeutralXMem := nx, NeutralYMem := ny);
home(DeadmanArmed := joy.DeadmanArmed, JoystickDeflected := NOT joy.AtNeutralXY, JoystickPull := joy.AxisCmdY.DirectionPositive, JoystickPush := joy.AxisCmdY.DirectionNegative, BtnValidation := bench.Operator.JoyBtnRaw);
ASSERT_EQ(home.MachineHomingSeqStep, E_MachineHomingTxState.HX0_REPOS, 'N1/cycle : aucun HX1 par geste joystick'); ASSERT_FALSE(home.M3Locked, 'N1/cycle : aucun verrou homing parasite'); ASSERT_TRUE(home.MachineHomed, 'Reference conservee');
ADVANCE_TIME(10000000); bench(RawPosM1 := raw1, RawPosM2 := raw2);
joy(RawX := bench.Operator.JoyXRaw_ANA1, RawY := bench.Operator.JoyYRaw_ANA2, RawButton := bench.Operator.JoyBtnRaw, Cfg := cfg, NeutralXMem := nx, NeutralYMem := ny);
home(DeadmanArmed := joy.DeadmanArmed, JoystickDeflected := NOT joy.AtNeutralXY, JoystickPull := joy.AxisCmdY.DirectionPositive, JoystickPush := joy.AxisCmdY.DirectionNegative, BtnValidation := bench.Operator.JoyBtnRaw);
ASSERT_EQ(home.MachineHomingSeqStep, E_MachineHomingTxState.HX0_REPOS, 'N1/cycle : aucun HX1 par geste joystick'); ASSERT_FALSE(home.M3Locked, 'N1/cycle : aucun verrou homing parasite'); ASSERT_TRUE(home.MachineHomed, 'Reference conservee');
END_TEST
